(* IEC 61131-3 sources: daoli-st-library/DL_Base (part 4) *)

(* ---- FC_DL_BitCountTransitions.st ---- *)
(*==============================================================================
 * 名称 : FC_DL_BitCountTransitions —— WORD 相邻位跳变统计（总跳变 / 上升 / 下降）
 * 分类 / 前缀 / 版本 : DL_Base / FC_DL_ / 1.0.0
 * 溯源 : 开源语义参考（OSCAT/AixOCAT 族，MIT）或 clean-room IEC 实现，未复制源码
 * 平台 : 纯 IEC 61131-3
 * 功能说明 : 单趟扫描 WORD 的 15 对相邻位（bit i-1 → bit i，i=1..15），统计
 *            跳变总次数并分解为上升（0→1）与下降（1→0）计数；恒有
 *            nRise + nFall = 返回值（调用方可据此自证）。
 *            边界处理：全 0 / 全 1 输入无跳变，三项全 0，属合法结果。
 * 错误码 : 无故障路径（全值域合法的纯统计），eErr 恒 0，bValid 恒 TRUE；
 *          16#0001_1A07 为本件预留码位，当前实现不发出
 * 状态机 : R6 标注 N/A（纯函数无顺序状态，以本节替代 ELSE 兜底）
 * 红线 : R1/R2/R3 ✓ 零全局/零IO/纯IEC ｜ R4 ✓ 移位量≤15 ｜ R10 ✓ 标准转换 ｜ R11 ✓ 分号收尾 ｜ R15 ✓ 无保留字撞名
 * 修订记录 : 2026-11-23 v1.0.0 首次入库（R76）
 *============================================================================*)
FUNCTION FC_DL_BitCountTransitions : INT
VAR_INPUT
    wWord : WORD;      // 待统计的输入字 [位域] / input word to be analyzed
END_VAR
VAR_OUTPUT
    nRise : INT;       // 0→1 上升跳变次数 [次] / number of rising transitions
    nFall : INT;       // 1→0 下降跳变次数 [次] / number of falling transitions
    eErr  : UDINT;     // 故障码，0=正常（本件无故障路径）/ error code, 0=ok (no fault path)
    bError: BOOL;      // 故障标志，恒 FALSE / error flag, always FALSE
    bValid: BOOL;      // TRUE=三项计数可用，恒 TRUE / TRUE when counts are usable
END_VAR
VAR
    _i     : INT;      // 位对扫描游标（取 bit i 与 bit i-1）[位] / pair scan cursor
    _wBit  : WORD;     // 当前位单比特掩码 [位域] / single-bit mask of current bit
    _wPrev : WORD;     // 前一位单比特掩码 [位域] / single-bit mask of previous bit
    _xCur  : BOOL;     // 当前位电平 / level of current bit
    _xPrev : BOOL;     // 前一位电平 / level of previous bit
END_VAR

FC_DL_BitCountTransitions := 0;              // 返回值（总跳变）预设 0 / preset total to zero
nRise := 0;                                  // 上升计数清零 / clear rise count
nFall := 0;                                  // 下降计数清零 / clear fall count
eErr  := 16#0000_0000;                       // 故障码清零 / clear error code
bError:= FALSE;                              // 故障标志清零 / clear error flag
bValid:= TRUE;                               // 本件全值域合法，恒可用 / always valid

FOR _i := 1 TO 15 DO                         // 扫描 15 对相邻位 / scan the 15 adjacent pairs
    _wBit  := SHL(WORD#16#0001, _i);         // 当前位掩码（_i≤15 安全）/ mask of current bit
    _wPrev := SHL(WORD#16#0001, _i - 1);     // 前一位掩码（i-1≥0 安全）/ mask of previous bit
    _xCur  := (wWord AND _wBit)  <> WORD#16#0000;    // 取当前位电平 / sample current bit
    _xPrev := (wWord AND _wPrev) <> WORD#16#0000;    // 取前一位电平 / sample previous bit
    IF _xCur AND (NOT _xPrev) THEN           // 0→1 上升沿 / rising transition
        nRise := nRise + 1;                  // 上升计数加一 / bump rise count
    END_IF
    IF (NOT _xCur) AND _xPrev THEN           // 1→0 下降沿 / falling transition
        nFall := nFall + 1;                  // 下降计数加一 / bump fall count
    END_IF
END_FOR

FC_DL_BitCountTransitions := nRise + nFall;  // 恒等式：总跳变 = 上升 + 下降 / invariant: total = rise + fall

END_FUNCTION

(* ---- FC_DL_BitFieldExtractLword.st ---- *)
(*
  ==================================================================
  组件名 Component  : FC_DL_BitFieldExtractLword
  分类   Category   : DL_Base
  复杂度 Complexity  : 中
  版本   Version    : 1.0.0
  功能   Purpose    : LWORD 单字段提取（起始位 + 宽度 → 右对齐字段值）。全程零
                      64 位移位：先拆高低两个 DWORD 半区，再在半区内做 <=31 位的
                      移位与常量掩码，跨半区时用 DWORD_TO_LWORD 升位拼接。
  来源   Source     : t2-1-lgf-bitlogic（LGF BitLogic 位域提取族 64 位变体）
  溯源   Origin     : 位域提取属公开位运算语义，clean-room 自研实现，未复制 LGF
                      或任何厂商私有库源码。
  平台   Platform   : 纯 IEC 61131-3（AND / OR / SHR / SHL 只作用在 DWORD 域，
                      移位量恒 <32；LWORD 域只出现 AND 与整除），三平台通用
  分工声明 Split     : 与 FC_DL_BitFieldExtract（32 位属主）互引——后者管 DWORD
                      域单字提取；本件为 LWORD 域半区拆分版，不重声明既有位域类型。
  作者   Author     : 道莅代码库 · PLC 编程专家（R60）
  ------------------------------------------------------------------
  边界 Boundary     :
                      一 全程零 64 位移位：高 32 位以「整除 2^32 再 LWORD_TO_DWORD」
                         取得（LWORD 域只做 AND 与整除，不做移位），半区内移位量
                         经 MOD 32 归一后恒在 0..31（R48）；
                      二 宽度 32 的掩码走常量 16#FFFF_FFFF，禁写 SHL(x, 32)；
                      三 非 32 对齐下「宽 64 跨两字」在本实现物理不可达（宽 64 只
                         能起始于位 0），此偏离显式声明：start + width > 64 时主动
                         收窄宽度并置截断信息级码，不静默出半个字段；
                      四 非法域：宽度为 0 或起始位 > 63 判故障级码，输出 0 且 bErr；
                      五 无状态纯函数：局部量一律段 1 显式预置（R254）。
  错误码   Codes    :
    16#0001_0616【故障级】字段域非法（宽度 0 或起始位 >63），输出 0
    16#0001_0617【信息级】字段越出 64 位容器，宽度已收窄（bTrunc 同步置位）
  验收   Acceptance :
    算法已证（脚本）：未跑 ｜ 编译器已证（三平台）：未跑
    V1 src=16#FFFF_FFFF_FFFF_FFFF、start=60、width=4 → 字段 16#F，bTrunc=FALSE
    V2 src=16#1234_5678_9ABC_DEF0、start=28、width=8 → 字段 16#BC（跨半区）
    V3 src 任意、start=62、width=8 → 宽度收窄为 2、bTrunc=TRUE、码 0617
    V4 width=0 → bErr=TRUE、码 0616、字段 0
  修订记录 Revision  :
    2026-11-21  v1.0.0  R60 首版（批 2 · 序号 5）
  ==================================================================
*)
FUNCTION FC_DL_BitFieldExtractLword : LWORD
VAR_INPUT
    uSrc   : LWORD; // 源字 [位串] / the source word
    uStart : UINT;  // 字段起始位号 [位]，合法域 0..63 / the field start bit, legal from zero to sixty three
    uWidth : UINT;  // 字段宽度 [位]，合法域 1..64 / the field width, legal from one to sixty four
END_VAR
VAR_OUTPUT
    bTrunc : BOOL;  // 宽度被收窄（越出容器）[-] / the width was narrowed at the container edge
    bErr   : BOOL;  // 域非法标志 [-] / the illegal domain flag
    eErr   : UDINT; // 错误码，0 = 正常 / the error code, zero is ok
    bError : BOOL;  // 错误标志，eErr 非 0 时为真 / the error flag, true when eErr is nonzero
END_VAR
VAR
    dwLow    : DWORD; // 源字低半区 [位串] / the low half of the source
    dwHigh   : DWORD; // 源字高半区 [位串] / the high half of the source
    dwMask   : DWORD; // 半区内字段掩码 [位串] / the field mask inside a half
    dwMaskHi : DWORD; // 跨半区时高半区剩余宽度掩码 [位串] / the remaining width mask on the high half
    dwPart1  : DWORD; // 跨半区低位片段 [位串] / the low fragment of a cross half field
    dwPart2  : DWORD; // 跨半区高位片段 [位串] / the high fragment of a cross half field
    nStart   : UINT;  // 归一后的起始位号 [位] / the normalised start bit
    nWidth   : UINT;  // 归一（收窄）后的宽度 [位] / the normalised width
    nLowW    : UINT;  // 跨半区时低半区可容纳宽度 [位] / the width the low half can hold
    nShift   : UINT;  // 半区内移位量 [位]，恒 0..31 / the shift amount inside a half, always zero through thirty one
END_VAR
VAR CONSTANT
    DL_BFE_32    : UINT := 32;                      // 半区位宽 [位] / the half width
    DL_BFE_ALL   : DWORD := 16#FFFF_FFFF;           // 32 位全一掩码（禁用 SHL(x, 32)）/ the full thirty two bit mask
    DL_BFE_2P32  : LWORD := 16#0000_0001_0000_0000; // 2 的 32 次幂，用于取高半区（LWORD 域整除，不做移位）/ two to the thirty second, used to take the high half by division
END_VAR

// 段 1｜返回值与错误状态预置安全值（四段式第一段，R45）+ 局部量显式预置（R254）/ segment 1, the preset of the return, the codes and the local guards
FC_DL_BitFieldExtractLword := 16#0000_0000_0000_0000; // 返回值预置零 / preset the return to zero
bTrunc := FALSE; // 截断标志预置假 / preset the truncation flag false
bErr := FALSE; // 域非法标志预置假 / preset the domain fault flag false
eErr := 16#0000_0000; // 错误码预置正常 / preset the code to ok
bError := FALSE; // 错误标志预置假 / preset the error flag false
nStart := 0; // 起始位预置零 / preset the start bit zero
nWidth := 0; // 宽度预置零 / preset the width zero
nLowW := 0; // 低半区宽度预置零 / preset the low half width zero
nShift := 0; // 移位量预置零 / preset the shift amount zero
dwMask := 16#0000_0000; // 掩码预置零 / preset the mask zero
dwMaskHi := 16#0000_0000; // 高位掩码预置零 / preset the high mask zero
dwPart1 := 16#0000_0000; // 低位片段预置零 / preset the low fragment zero
dwPart2 := 16#0000_0000; // 高位片段预置零 / preset the high fragment zero

// 段 2｜域闸（下界早退 + 上界钳位，边界三）/ segment 2, the domain gate with the early return and the narrowing
IF (uWidth < 1) OR (uStart > 63) THEN // 宽度为零或起始位越域 / a zero width or a start beyond the container
    bErr := TRUE; // 置域非法标志 / raise the domain fault flag
    eErr := 16#0001_0616; // 故障级：字段域非法 / fault grade, the field domain is illegal
    bError := TRUE; // 置错误标志（R45 配对）/ raise the error flag, paired with the fault code
    RETURN; // 早退：返回值保持零 / early return with the field zero
END_IF
nStart := uStart; // 域内接管起始位 / take the start bit inside the domain
nWidth := uWidth; // 域内接管宽度 / take the width inside the domain
IF (UINT_TO_UDINT(nStart) + UINT_TO_UDINT(nWidth)) > 64 THEN // 越出 64 位容器 / beyond the sixty four bit container
    nWidth := 64 - nStart; // 主动收窄到容器边界（边界三偏离声明）/ narrow to the container edge with the declared deviation
    bTrunc := TRUE; // 置截断标志 / raise the truncation flag
    eErr := 16#0001_0617; // 信息级：宽度已收窄 / informational, the width narrowed
    bError := TRUE; // 置错误标志 / raise the error flag
END_IF

// 段 3｜半区拆分（零 64 位移位，边界一）：低半区截断取，高半区整除取 / segment 3, the half split with no sixty four bit shift
dwLow := LWORD_TO_DWORD(uSrc); // 低半区：截断取低 32 位 / the low half by truncation
dwHigh := LWORD_TO_DWORD(uSrc / DL_BFE_2P32); // 高半区：整除 2^32 后取低 32 位 / the high half by the division

// 段 4｜字段提取与跨半区拼接（掩码先于移位构造，移位量恒 <32）/ segment 4, the extraction and the cross half splice
IF (nWidth = 32) THEN // 宽 32：常量全一掩码（禁 SHL(x, 32)）/ a full half width uses the constant mask
    dwMask := DL_BFE_ALL; // 常量掩码 / the constant mask
ELSE // 宽 1..31：SHL(1, nWidth) - 1，移位量最大 31 结构性安全 / widths one through thirty one
    dwMask := SHL(DWORD#1, nWidth) - DWORD#1; // 低位起的 nWidth 个一并 / the nWidth low bits set
END_IF
IF nStart >= DL_BFE_32 THEN // 字段整段落在高半区 / the field lies entirely in the high half
    nShift := nStart - DL_BFE_32; // 半区内移位量 0..31 / the shift inside the half, zero through thirty one
    FC_DL_BitFieldExtractLword := DWORD_TO_LWORD(SHR(dwHigh AND dwMask, nShift)); // 高半区提取后升位 / extract from the high half then widen
ELSIF (UINT_TO_UDINT(nStart) + UINT_TO_UDINT(nWidth)) <= 32 THEN // 字段整段落在低半区 / the field lies entirely in the low half
    nShift := nStart; // 半区内移位量 0..31 / the shift inside the half, zero through thirty one
    FC_DL_BitFieldExtractLword := DWORD_TO_LWORD(SHR(dwLow AND dwMask, nShift)); // 低半区提取后升位 / extract from the low half then widen
ELSE // 跨半区：低片段 + 高片段移位拼接（nStart 必在 1..31）/ a cross half field, both fragments spliced
    nLowW := 32 - nStart; // 低半区可容纳宽度 1..31 / the width the low half holds, one through thirty one
    IF nLowW >= 32 THEN // 结构性不可达（nStart ≥ 1 恒真），显式兜底防掩码移位越界 / structurally unreachable, kept as an explicit guard
        nLowW := 31; // 兜底收窄到 31 位 / narrow to thirty one bits
    END_IF
    dwPart1 := SHR(dwLow AND (SHL(DWORD#1, nLowW) - DWORD#1), nStart); // 低片段右移到最低位 / shift the low fragment down to bit zero
    dwMaskHi := SHL(DWORD#1, nWidth - nLowW) - DWORD#1; // 高半区剩余宽度掩码 / the remaining width mask on the high half
    dwPart2 := SHL(dwHigh AND dwMaskHi, nLowW); // 高片段左移到低片段之上（移位量 1..31）/ shift the high fragment above the low one
    FC_DL_BitFieldExtractLword := DWORD_TO_LWORD(dwPart1 OR dwPart2); // 两片段拼合后升位 / splice then widen
END_IF

// 段 5｜结果复检：字段宽度上界自证（nWidth ≤ 64，拼接已按半区完成，无溢出路径）/ segment 5, the result recheck
IF bTrunc AND (nWidth >= 1) THEN // 收窄后仍为合法宽度 / the narrowed width is still legal
    eErr := 16#0001_0617; // 信息级：宽度已收窄（回放，防段 4 覆盖）/ informational, the width narrowed, replayed against the overwrite
END_IF
END_FUNCTION

(* ---- FC_DL_BitFillLowestZero.st ---- *)
(*==============================================================================
 * 名称 : FC_DL_BitFillLowestZero —— 最低 0 位置 1（DWORD），输出该位位号
 * 分类 / 前缀 / 版本 : DL_Base / FC_DL_ / 1.0.0
 * 溯源 : 开源语义参考（OSCAT/AixOCAT 族，MIT）或 clean-room IEC 实现，未复制源码
 * 平台 : 纯 IEC 61131-3
 * 功能说明 : 把输入 DWORD 中最低的 0 位置 1 后返回（即 dwIn OR 单比特隔离值），
 *            并给出该位位号 nPos。常用于资源位图分配（找空位并占用）。
 *            边界处理：输入全 1 时无 0 位可填，原值返回、nPos=-1、bValid=FALSE
 *            并置 eErr（返回值虽为原值，但语义上未发生分配）。
 * 错误码 : 16#0001_1A08 = 输入全 1，无 0 位可填
 *          eErr=0 且 bValid=TRUE 表示已完成填位且 nPos 有效
 * 状态机 : R6 标注 N/A（纯函数无顺序状态，以本节替代 ELSE 兜底）
 * 红线 : R1/R2/R3 ✓ 零全局/零IO/纯IEC ｜ R4 ✓ 移位量≤31 ｜ R10 ✓ 标准转换 ｜ R11 ✓ 分号收尾 ｜ R15 ✓ 无保留字撞名
 * 修订记录 : 2026-11-23 v1.0.0 首次入库（R76）
 *============================================================================*)
FUNCTION FC_DL_BitFillLowestZero : DWORD
VAR_INPUT
    dwIn : DWORD;      // 输入位图 [位域] / input bitmap dword
END_VAR
VAR_OUTPUT
    nPos   : INT;      // 被填 1 的最低 0 位位号，全 1 时为 -1 [位] / bit index filled, -1 if none
    eErr   : UDINT;    // 故障码，0=正常，1A08=全 1 无空位 / error code, 0=ok, 1A08=all-ones input
    bError : BOOL;     // TRUE=本件发生故障 / TRUE when fault occurred
    bValid : BOOL;     // TRUE=填位成功且 nPos 有效 / TRUE when fill succeeded and nPos valid
END_VAR
VAR
    _dwNot  : DWORD;   // 输入按位取反（0 位变 1 位）/ inverted input (zeros become ones)
    _dwIso  : DWORD;   // 最低 0 位的单比特隔离值 [位域] / isolated lowest zero bit
    _i      : INT;     // 位扫描游标 [位] / bit scan cursor
    _dwW    : DWORD;   // 单比特游走值 [位域] / single-bit walker
    _xHit   : BOOL;    // 命中标志 / found flag
END_VAR

nPos := -1;                                  // 位号预设 -1（未命中语义）/ preset position to -1
eErr   := 16#0000_0000;                      // 故障码清零 / clear error code
bError := FALSE;                             // 故障标志清零 / clear error flag
bValid := TRUE;                              // 预设输出可用 / preset valid flag

_dwNot := NOT dwIn;                          // 取反后 0 位变 1 位 / invert so zeros become ones
IF _dwNot = DWORD#16#0000_0000 THEN          // 全 1：无 0 位可填 / all ones: nothing to fill
    eErr   := 16#0001_1A08;                  // 置全 1 故障码 / set all-ones code
    bError := TRUE;                          // 置故障标志 / set error flag
    bValid := FALSE;                         // nPos 不可用 / position not usable
    FC_DL_BitFillLowestZero := dwIn;         // 原值返回 / return input unchanged
    RETURN;                                  // 提前收口 / early exit
END_IF

_dwIso := _dwNot AND (NOT (_dwNot - DWORD#16#0000_0001));    // 隔离最低 0 位（同最低 1 位法）/ isolate lowest zero bit
_xHit  := FALSE;                             // 命中标志清零 / clear found flag
FOR _i := 0 TO 31 DO                         // 从低位找第一个命中 / scan low to high for first hit
    _dwW := SHL(DWORD#16#0000_0001, _i);     // 当前位单比特掩码（_i≤31 安全）/ single-bit mask
    IF (NOT _xHit) AND ((_dwIso AND _dwW) <> DWORD#16#0000_0000) THEN    // 首个命中即停扫 / stop at first hit
        nPos  := _i;                         // 回写位号 / write back bit index
        _xHit := TRUE;                       // 置命中标志 / set found flag
    END_IF
END_FOR

FC_DL_BitFillLowestZero := dwIn OR _dwIso;   // 填 1 后返回 / return with the bit filled

END_FUNCTION

(* ---- FC_DL_BitGet.st ---- *)
(*==============================================================================
 * 组件名称 (Component)  : FC_DL_BitGet
 * 所属子库 (Sublibrary) : DL_Base
 * 当前版本 (Version)    : 1.0.0
 * 兼容性   (Platform)   : CODESYS 3.5 / TwinCAT 3 / 汇川 InoProShop / Machine Expert
 *                         仅用标准 SHR / AND 运算，无任何厂商位访问语法
 * 功能描述 (Function)   : 从 32 位状态字中安全提取指定位（Hamming 单位提取）。
 *                         位索引合法域 0..31（0 = LSB）。越界时"先判后算"，
 *                         立即返回 FALSE 并输出 16#0001_0001，绝不把越界移位量
 *                         交给 SHL/SHR 去执行（越界移位在各平台行为不一致，是
 *                         跨平台移植的经典暗坑）。
 * 开源溯源 (Origin)     : 原创实现。位序约定遵循 IEC 61131-3 对位串类型
 *                         "第 0 位为最低有效位"的规定。
 * 依赖     (Depends)    : 无 DL_ 内部依赖；无标准库功能块依赖
 * 红线自检 (Redline)    : R1 ✓ 零全局变量表与外部变量引用 ｜ R2 ✓ 零物理 IO 地址直写
 *                         R3 ✓ 纯 IEC 61131-3（无厂商位访问方言）｜ R4 ✓ 越界先判后算 + 返回值兜底
 *                         R5 ✓ 全变量中英双语同行注释 ｜ R6 N/A（无状态机）｜ R7 N/A（无实例调用）
 * 修订历史 (Revision)   :
 *   2026-11-14  v1.0.0  首版入库（Phase 1 冷启动 · Level 0 批次）
 *============================================================================*)
FUNCTION FC_DL_BitGet : BOOL
VAR_INPUT
    uValue    : DWORD;    // 待检测的 32 位状态字 / Source 32-bit status word
    uBitIndex : USINT;    // 位序号，0 = LSB，合法域 0..31 / Bit index, 0 = LSB, valid range 0..31
END_VAR
VAR_OUTPUT
    bValid    : BOOL;     // 索引合法标志，FALSE 时返回值为保底 FALSE / Index valid flag, FALSE means result is a safe FALSE
    uErrorId  : UDINT;    // 故障码，0 = 无故障 / Error code, 0 = no error
END_VAR
VAR
    uWork     : UDINT;    // 提升到 UDINT 的工作副本，规避混合类型移位 / UDINT working copy to avoid mixed-type shifts
    uShift    : UDINT;    // 提升到 UDINT 的移位量 / Shift amount promoted to UDINT
END_VAR
VAR CONSTANT
    DL_BIT_INDEX_MAX : USINT := 31;  // 32 位字的最大合法位索引 / Max legal bit index of a 32-bit word
END_VAR

(*------------------------------------------------------------------------------
 * 段 1｜返回值与标志预置：任何异常路径下返回值必须确定
 *      Pre-set return value and flags: the result must be deterministic on every path
 *      部分平台函数返回值未赋值时残留上次调用值，故先给 FALSE（边界 B4）
 *-----------------------------------------------------------------------------*)
FC_DL_BitGet := FALSE;
bValid       := FALSE;
uErrorId     := 16#0000_0000;
uWork        := 16#0000_0000;

(*------------------------------------------------------------------------------
 * 段 2｜越界先判后算（边界 B1）：禁止先移位再校验
 *      Bounds check before any shift (boundary B1): never shift first and check later
 *      USINT 全域 0..255，凡 > 31 者均属非法移位量，统一按参数越界处理
 *-----------------------------------------------------------------------------*)
IF uBitIndex > DL_BIT_INDEX_MAX THEN
    uErrorId := 16#0001_0001;
    RETURN;
END_IF

(*------------------------------------------------------------------------------
 * 段 3｜位提取（边界 B2/B3）：统一提升到 UDINT 后移位，再显式掩码取最低位
 *      Bit extraction: promote to UDINT, shift, then mask the LSB explicitly
 *      禁止使用以点号直取单一位的厂商方言；禁止依赖"非零即真"的隐式布尔转换
 *-----------------------------------------------------------------------------*)
uWork  := DWORD_TO_UDINT(uValue);
uShift := USINT_TO_UDINT(uBitIndex);
uWork  := SHR(uWork, uShift);
uWork  := uWork AND 16#0000_0001;

IF uWork <> 16#0000_0000 THEN
    FC_DL_BitGet := TRUE;
END_IF

(* 校验通过：索引合法，结果可信 *)
(* Check passed: index is legal and the result is trustworthy *)
bValid := TRUE;
END_FUNCTION

(* ---- FC_DL_BitLowestSet.st ---- *)
(*==============================================================================
 * 名称 : FC_DL_BitLowestSet —— 最低置位位号与单比特隔离值（DWORD）
 * 分类 / 前缀 / 版本 : DL_Base / FC_DL_ / 1.0.0
 * 溯源 : 开源语义参考（OSCAT/AixOCAT 族，MIT）或 clean-room IEC 实现，未复制源码
 * 平台 : 纯 IEC 61131-3
 * 功能说明 : 返回输入 DWORD 中最低置位位的位号（0..31），并输出单比特隔离值
 *            dwIsolate = dwIn AND (NOT (dwIn - 1))（无符号回绕语义，等价于
 *            二进制补码的 x AND (-x)，仅保留最低的 1 位）。
 *            边界处理：dwIn 全 0 时无置位位，返回 -1、dwIsolate=0、bValid=FALSE
 *            并置 eErr（隔离值无效，调用方不得使用）。
 * 错误码 : 16#0001_1A05 = 输入全 0，无置位位可隔离
 *          eErr=0 且 bValid=TRUE 表示返回位号与隔离值均有效
 * 状态机 : R6 标注 N/A（纯函数无顺序状态，以本节替代 ELSE 兜底）
 * 红线 : R1/R2/R3 ✓ 零全局/零IO/纯IEC ｜ R4 ✓ 移位量≤31 ｜ R10 ✓ 标准转换 ｜ R11 ✓ 分号收尾 ｜ R15 ✓ 无保留字撞名
 * 修订记录 : 2026-11-23 v1.0.0 首次入库（R76）
 *============================================================================*)
FUNCTION FC_DL_BitLowestSet : INT
VAR_INPUT
    dwIn : DWORD;      // 待扫描的输入双字 [位域] / input dword to be scanned
END_VAR
VAR_OUTPUT
    dwIsolate : DWORD;    // 最低置位位的单比特隔离值 [位域] / isolated lowest set bit
    eErr      : UDINT;    // 故障码，0=正常，1A05=输入全 0 / error code, 0=ok, 1A05=all-zero input
    bError    : BOOL;     // TRUE=本件发生故障 / TRUE when fault occurred
    bValid    : BOOL;     // TRUE=返回位号与隔离值可用 / TRUE when outputs are usable
END_VAR
VAR
    _i    : INT;       // 位扫描游标 [位] / bit scan cursor
    _dwW  : DWORD;     // 单比特游走值 [位域] / single-bit walker
    _xHit : BOOL;      // 是否已找到最低置位位 / found flag for lowest set bit
END_VAR

FC_DL_BitLowestSet := -1;                    // 返回值预设 -1（未命中语义）/ preset return to -1
dwIsolate := DWORD#16#0000_0000;             // 隔离值预设全 0 / preset isolate to zero
eErr      := 16#0000_0000;                   // 故障码清零 / clear error code
bError    := FALSE;                          // 故障标志清零 / clear error flag
bValid    := TRUE;                           // 预设输出可用 / preset valid flag

IF dwIn = DWORD#16#0000_0000 THEN            // 输入全 0：无置位位 / all-zero input: no set bit
    eErr   := 16#0001_1A05;                  // 置全 0 故障码 / set all-zero code
    bError := TRUE;                          // 置故障标志 / set error flag
    bValid := FALSE;                         // 位号与隔离值均不可用 / outputs not usable
    RETURN;                                  // 返回 -1、隔离值 0 / return -1 with zero isolate
END_IF

dwIsolate := dwIn AND (NOT (dwIn - DWORD#16#0000_0001));    // 经典隔离式，仅留最低 1 位 / classic isolate of lowest set bit
_xHit := FALSE;                              // 命中标志清零 / clear found flag
FOR _i := 0 TO 31 DO                         // 从低位向高位找第一个 1 / scan low to high for first one
    _dwW := SHL(DWORD#16#0000_0001, _i);     // 当前位单比特掩码（_i≤31 安全）/ single-bit mask
    IF (NOT _xHit) AND ((dwIsolate AND _dwW) <> DWORD#16#0000_0000) THEN    // 首个命中即停扫 / stop at first hit
        FC_DL_BitLowestSet := _i;            // 回写最低置位位号 / write back lowest bit index
        _xHit := TRUE;                       // 置命中标志 / set found flag
    END_IF
END_FOR

END_FUNCTION

(* ---- FC_DL_BitMaskRange.st ---- *)
(*==============================================================================
 * 名称 : FC_DL_BitMaskRange —— 连续位区间掩码构造（bitLo..bitHi 置 1 的 DWORD 掩码）
 * 分类 / 前缀 / 版本 : DL_Base / FC_DL_ / 1.0.0
 * 溯源 : 开源语义参考（OSCAT/AixOCAT 族，MIT）或 clean-room IEC 实现，未复制源码
 * 平台 : 纯 IEC 61131-3
 * 功能说明 : 依入参位号 uLo..uHi 构造 DWORD 掩码，区间内各位置 1、其余为 0。
 *            边界处理：uLo/uHi 越界（<0 或 >31）先钳位到 [0,31] 再构造；
 *            钳位后 uLo>uHi（区间为空）返回 DWORD#0 并置 eErr 故障码。
 *            移位量恒 ≤31（<DWORD 位宽 32），结构性无越界移位。
 * 错误码 : 16#0001_1A01 = 钳位后位区间为空（uLo>uHi），掩码无意义
 *          eErr=0 且 bValid=TRUE 表示掩码有效；bValid=FALSE 时返回值勿用
 * 状态机 : R6 标注 N/A（纯函数无顺序状态，以本节替代 ELSE 兜底）
 * 红线 : R1/R2/R3 ✓ 零全局/零IO/纯IEC ｜ R4 ✓ 移位量≤31 ｜ R10 ✓ 标准转换 ｜ R11 ✓ 分号收尾 ｜ R15 ✓ 无保留字撞名
 * 修订记录 : 2026-11-23 v1.0.0 首次入库（R76）
 *============================================================================*)
FUNCTION FC_DL_BitMaskRange : DWORD
VAR_INPUT
    uLo : INT;     // 起始位号 0..31，越界自动钳位 [位] / low bit index, clamped into [0,31]
    uHi : INT;     // 结束位号 0..31，越界自动钳位 [位] / high bit index, clamped into [0,31]
END_VAR
VAR_OUTPUT
    eErr   : UDINT;    // 故障码，0=正常，1A01=区间为空 / error code, 0=ok, 1A01=empty range
    bError : BOOL;     // TRUE=本件发生参数级故障 / TRUE when parameter-level fault occurred
    bValid : BOOL;     // TRUE=返回值可用 / TRUE when return value is usable
END_VAR
VAR
    _nLo   : INT;      // 钳位后的起始位号 [位] / clamped low bit index
    _nHi   : INT;      // 钳位后的结束位号 [位] / clamped high bit index
    _i     : INT;      // 位扫描游标 [位] / bit scan cursor
    _dwBit : DWORD;    // 当前游标对应的单比特值 [位域] / single-bit walker value
END_VAR

FC_DL_BitMaskRange := DWORD#16#0000_0000;    // 返回值预设全 0 掩码 / preset return to zero mask
eErr   := 16#0000_0000;                      // 故障码清零 / clear error code
bError := FALSE;                             // 故障标志清零 / clear error flag
bValid := TRUE;                              // 预设输出可用 / preset valid flag

_nLo := uLo;                                 // 取入参起始位号 / take input low index
_nHi := uHi;                                 // 取入参结束位号 / take input high index
IF _nLo < 0 THEN _nLo := 0; END_IF           // 下界钳位 / clamp lower bound
IF _nLo > 31 THEN _nLo := 31; END_IF         // 上界钳位 / clamp upper bound
IF _nHi < 0 THEN _nHi := 0; END_IF           // 下界钳位 / clamp lower bound
IF _nHi > 31 THEN _nHi := 31; END_IF         // 上界钳位 / clamp upper bound

IF _nLo > _nHi THEN                          // 钳位后区间为空 / empty range after clamping
    eErr   := 16#0001_1A01;                  // 置区间为空故障码 / set empty-range code
    bError := TRUE;                          // 置故障标志 / set error flag
    bValid := FALSE;                         // 返回值不可用 / return value not usable
    RETURN;                                  // 返回值保持全 0 掩码 / return stays zero mask
END_IF

_dwBit := SHL(DWORD#16#0000_0001, _nLo);     // 单比特走到起始位（_nLo≤31 安全）/ walk bit to start
FOR _i := _nLo TO _nHi DO                    // 逐位置 1 / set bits one by one
    FC_DL_BitMaskRange := FC_DL_BitMaskRange OR _dwBit;    // 并入当前位 / merge current bit
    _dwBit := SHL(_dwBit, 1);                // 单比特左移一位，循环内 _i<_nHi≤31 安全 / shift walker left
END_FOR

END_FUNCTION

(* ---- FC_DL_BitReverse16.st ---- *)
(*==============================================================================
 * 名称 : FC_DL_BitReverse16 —— WORD 位序完全反转（bit0↔bit15 镜像）
 * 分类 / 前缀 / 版本 : DL_Base / FC_DL_ / 1.0.0
 * 溯源 : 开源语义参考（OSCAT/AixOCAT 族，MIT）或 clean-room IEC 实现，未复制源码
 * 平台 : 纯 IEC 61131-3
 * 功能说明 : 将 WORD 的 16 个位按镜像序重排后返回（第 i 位映射到第 15-i 位）。
 *            边界处理：全 0 / 全 1 / 回文位型（如 16#8081）均原值返回，属合法结果；
 *            循环固定 16 次，无越界移位（i 与 15-i 均 ≤15 < 16 位宽）。
 * 错误码 : 无故障路径（全值域合法的纯变换），eErr 恒 0，bValid 恒 TRUE；
 *          16#0001_1A03 为本件预留码位，当前实现不发出
 * 状态机 : R6 标注 N/A（纯函数无顺序状态，以本节替代 ELSE 兜底）
 * 红线 : R1/R2/R3 ✓ 零全局/零IO/纯IEC ｜ R4 ✓ 移位量≤15 ｜ R10 ✓ 标准转换 ｜ R11 ✓ 分号收尾 ｜ R15 ✓ 无保留字撞名
 * 修订记录 : 2026-11-23 v1.0.0 首次入库（R76）
 *============================================================================*)
FUNCTION FC_DL_BitReverse16 : WORD
VAR_INPUT
    wIn : WORD;        // 待反转的输入字 [位域] / input word to be bit-reversed
END_VAR
VAR_OUTPUT
    eErr   : UDINT;    // 故障码，0=正常（本件无故障路径）/ error code, 0=ok (no fault path)
    bError : BOOL;     // 故障标志，恒 FALSE / error flag, always FALSE
    bValid : BOOL;     // TRUE=返回值可用，恒 TRUE / TRUE when return value is usable
END_VAR
VAR
    _i     : INT;      // 位扫描游标 [位] / bit scan cursor
    _wBit  : WORD;     // 当前读出位对应的单比特值 [位域] / single-bit walker for read side
END_VAR

FC_DL_BitReverse16 := WORD#16#0000;          // 返回值预设全 0 / preset return to zero
eErr   := 16#0000_0000;                      // 故障码清零 / clear error code
bError := FALSE;                             // 故障标志清零 / clear error flag
bValid := TRUE;                              // 本件全值域合法，恒可用 / always valid

FOR _i := 0 TO 15 DO                         // 逐位镜像搬运 / mirror bits one by one
    _wBit := SHL(WORD#16#0001, _i);          // 读侧单比特（_i≤15 安全）/ single bit on read side
    IF (wIn AND _wBit) <> WORD#16#0000 THEN  // 源位为 1 才搬运 / copy only when source bit set
        FC_DL_BitReverse16 := FC_DL_BitReverse16 OR SHL(WORD#16#0001, 15 - _i);    // 写入镜像位（15-_i≤15 安全）/ set mirrored bit
    END_IF
END_FOR

END_FUNCTION

(* ---- FC_DL_BitReverse8.st ---- *)
(*==============================================================================
 * 名称 : FC_DL_BitReverse8 —— BYTE 位序完全反转（bit0↔bit7 镜像）
 * 分类 / 前缀 / 版本 : DL_Base / FC_DL_ / 1.0.0
 * 溯源 : 开源语义参考（OSCAT/AixOCAT 族，MIT）或 clean-room IEC 实现，未复制源码
 * 平台 : 纯 IEC 61131-3
 * 功能说明 : 将 BYTE 的 8 个位按镜像序重排后返回（第 i 位映射到第 7-i 位）。
 *            边界处理：全 0 / 全 1 / 回文位型（如 16#18）均原值返回，属合法结果；
 *            循环固定 8 次，无越界移位（i 与 7-i 均 ≤7 < 8 位宽）。
 * 错误码 : 无故障路径（全值域合法的纯变换），eErr 恒 0，bValid 恒 TRUE；
 *          16#0001_1A02 为本件预留码位，当前实现不发出
 * 状态机 : R6 标注 N/A（纯函数无顺序状态，以本节替代 ELSE 兜底）
 * 红线 : R1/R2/R3 ✓ 零全局/零IO/纯IEC ｜ R4 ✓ 移位量≤7 ｜ R10 ✓ 标准转换 ｜ R11 ✓ 分号收尾 ｜ R15 ✓ 无保留字撞名
 * 修订记录 : 2026-11-23 v1.0.0 首次入库（R76）
 *============================================================================*)
FUNCTION FC_DL_BitReverse8 : BYTE
VAR_INPUT
    byIn : BYTE;       // 待反转的输入字节 [位域] / input byte to be bit-reversed
END_VAR
VAR_OUTPUT
    eErr   : UDINT;    // 故障码，0=正常（本件无故障路径）/ error code, 0=ok (no fault path)
    bError : BOOL;     // 故障标志，恒 FALSE / error flag, always FALSE
    bValid : BOOL;     // TRUE=返回值可用，恒 TRUE / TRUE when return value is usable
END_VAR
VAR
    _i     : INT;      // 位扫描游标 [位] / bit scan cursor
    _dwBit : BYTE;     // 当前读出位对应的单比特值 [位域] / single-bit walker for read side
END_VAR

FC_DL_BitReverse8 := BYTE#16#00;             // 返回值预设全 0 / preset return to zero
eErr   := 16#0000_0000;                      // 故障码清零 / clear error code
bError := FALSE;                             // 故障标志清零 / clear error flag
bValid := TRUE;                              // 本件全值域合法，恒可用 / always valid

FOR _i := 0 TO 7 DO                          // 逐位镜像搬运 / mirror bits one by one
    _dwBit := SHL(BYTE#16#01, _i);           // 读侧单比特（_i≤7 安全）/ single bit on read side
    IF (byIn AND _dwBit) <> BYTE#16#00 THEN  // 源位为 1 才搬运 / copy only when source bit set
        FC_DL_BitReverse8 := FC_DL_BitReverse8 OR SHL(BYTE#16#01, 7 - _i);    // 写入镜像位（7-_i≤7 安全）/ set mirrored bit
    END_IF
END_FOR

END_FUNCTION

(* ---- FC_DL_BitRunLength.st ---- *)
(*==============================================================================
 * 名称 : FC_DL_BitRunLength —— WORD 最长连续 1 游程长度与起始位号
 * 分类 / 前缀 / 版本 : DL_Base / FC_DL_ / 1.0.0
 * 溯源 : 开源语义参考（OSCAT/AixOCAT 族，MIT）或 clean-room IEC 实现，未复制源码
 * 平台 : 纯 IEC 61131-3
 * 功能说明 : 单趟扫描 WORD 的 16 个位，返回最长连续 1 的游程长度（0..16），
 *            并给出该游程的起始位号 nStart（0..15）。多条等长游程取最低起始位。
 *            边界处理：无任何 1 位时返回 0 且 nStart=-1（合法结果，非故障，
 *            bValid 保持 TRUE）；游程到字尾截断同样按已计长度参与比较。
 * 错误码 : 无故障路径（全值域合法的纯统计），eErr 恒 0，bValid 恒 TRUE；
 *          16#0001_1A04 为本件预留码位，当前实现不发出
 * 状态机 : R6 标注 N/A（纯函数无顺序状态，以本节替代 ELSE 兜底）
 * 红线 : R1/R2/R3 ✓ 零全局/零IO/纯IEC ｜ R4 ✓ 移位量≤15 ｜ R10 ✓ 标准转换 ｜ R11 ✓ 分号收尾 ｜ R15 ✓ 无保留字撞名
 * 修订记录 : 2026-11-23 v1.0.0 首次入库（R76）
 *============================================================================*)
FUNCTION FC_DL_BitRunLength : INT
VAR_INPUT
    wWord : WORD;      // 待扫描的输入字 [位域] / input word to be scanned
END_VAR
VAR_OUTPUT
    nStart : INT;      // 最长游程起始位号，无 1 时为 -1 [位] / start bit of longest run, -1 if none
    eErr   : UDINT;    // 故障码，0=正常（本件无故障路径）/ error code, 0=ok (no fault path)
    bError : BOOL;     // 故障标志，恒 FALSE / error flag, always FALSE
    bValid : BOOL;     // TRUE=返回值可用，恒 TRUE / TRUE when return value is usable
END_VAR
VAR
    _i        : INT;       // 位扫描游标 [位] / bit scan cursor
    _nCur     : INT;       // 当前游程长度 [位] / current run length
    _nCurSt   : INT;       // 当前游程起始位号 [位] / current run start bit
    _nBest    : INT;       // 已发现的最长游程长度 [位] / best run length so far
    _nBestSt  : INT;       // 已发现的最长游程起始位号 [位] / best run start bit so far
    _wBit     : WORD;      // 当前位单比特掩码 [位域] / single-bit mask of current position
    _xBit     : BOOL;      // 当前位电平 / level of current bit
END_VAR

FC_DL_BitRunLength := 0;                     // 返回值预设 0 / preset return to zero
nStart := -1;                                // 起始位预设 -1（无 1 语义）/ preset start to -1
eErr   := 16#0000_0000;                      // 故障码清零 / clear error code
bError := FALSE;                             // 故障标志清零 / clear error flag
bValid := TRUE;                              // 本件全值域合法，恒可用 / always valid

_nBest  := 0;                                // 最长游程清零 / clear best length
_nBestSt := -1;                              // 最长游程起始清零 / clear best start
_nCur   := 0;                                // 当前游程清零 / clear current length
_nCurSt := 0;                                // 当前游程起始清零 / clear current start

FOR _i := 0 TO 15 DO                         // 单趟从低位到高位扫描 / single low-to-high pass
    _wBit := SHL(WORD#16#0001, _i);          // 当前位单比特掩码（_i≤15 安全）/ single-bit mask
    _xBit := (wWord AND _wBit) <> WORD#16#0000;    // 取当前位电平 / sample current bit
    IF _xBit THEN                            // 位为 1：游程延续或新开 / bit set: extend or open run
        IF _nCur = 0 THEN
            _nCurSt := _i;                   // 新游程序幕，记起始位 / new run starts here
        END_IF
        _nCur := _nCur + 1;                  // 游程长度加一 / extend run length
        IF _nCur > _nBest THEN               // 严格大于保证等长取最低起始位 / strict gt keeps lowest start on ties
            _nBest   := _nCur;               // 刷新最长游程 / refresh best length
            _nBestSt := _nCurSt;             // 刷新最长游程起始位 / refresh best start bit
        END_IF
    ELSE                                     // 位为 0：当前游程终结 / bit clear: current run ends
        _nCur := 0;                          // 游程长度归零 / reset current length
    END_IF
END_FOR

FC_DL_BitRunLength := _nBest;                // 回写最长游程长度 / write back best length
nStart := _nBestSt;                          // 回写起始位号（无 1 时保持 -1）/ write back start bit

END_FUNCTION

(* ---- FC_DL_BitScanLword.st ---- *)
(*
  ==================================================================
  组件名 Component  : FC_DL_BitScanLword
  分类   Category   : DL_Base
  前缀   Naming     : FC_DL_ ｜ b/n/u/f/t/e/st 类型前缀制（R265）
  复杂度 Complexity  : 低
  版本   Version    : 1.0.0
  功能   Purpose    : LWORD 最低/最高置位索引扫描（uIdx + bFound 双出口）。
  来源   Source     : self-std（IEC 标准位操作语义自研包装）
  平台   Platform   : 纯 IEC 61131-3（FOR / AND / SHR / SHL / 比较），三平台通用
  分工声明 Split     : 与 FC_DL_ReverseBitsLword（位序反转属主）分工——本件只做
                      置位索引定位，不改位序；方向由 bHighFirst 选择，不设两个 POU。
  作者   Author     : 道莅代码库 · PLC 编程专家（R61）
  归属 Ownership     : 本件无 TYPE 声明；引用件类型全部 IEC 标准原生。
  ------------------------------------------------------------------
  边界 Boundary     :
                      一 全零输入：bFound = FALSE 且 uIdx = 0（不泄 -1，不泄哨兵），
                         置信息级码（R90 反证：bFound 只表达「有命中」，无法区分
                         「扫描过且全零」与「未扫」，码位补足该可观测性）；
                      二 扫描循环有界恰好 64 次（禁 WHILE 裸循环，防死锁纪律）；
                      三 方向选择：bHighFirst = FALSE 自低位向高位扫（首命中即
                         最低置位），TRUE 自高位向低位扫（首命中即最高置位）；
                      四 无状态纯函数：局部量段 1 显式预置（R254）。
  错误码   Codes    :
    16#0001_0641【信息级】全零输入零命中（bFound = FALSE，uIdx = 0）
  验收   Acceptance :
    算法已证（脚本）：未跑 ｜ 编译器已证（三平台）：未跑
    V1 uSrc=16#0000_0000_0000_0100、bHighFirst=FALSE → uIdx=8、bFound=TRUE
    V2 uSrc=16#0000_0000_0000_0100、bHighFirst=TRUE → uIdx=8（单置位两向同值）
    V3 uSrc=16#0000_0000_0000_0105、bHighFirst=TRUE → uIdx=8
    V4 uSrc=0 → bFound=FALSE、uIdx=0、码 0641
  修订记录 Revision  :
    2026-11-21  v1.0.0  R61 首版（批 1 · 序号 2）
  ==================================================================
*)
FUNCTION FC_DL_BitScanLword : BOOL
VAR_IN_OUT
    uSrc : LWORD; // 待扫描源字 [位图] / the source word to scan
END_VAR
VAR_INPUT
    bHighFirst : BOOL; // 方向开关：TRUE 自高位向低位扫 / the direction switch, true scans from the high end
END_VAR
VAR_OUTPUT
    uIdx   : UDINT; // 首命中置位索引 [位]，零命中时为 0 / the first hit bit index, zero on a miss
    bFound : BOOL;  // 是否存在置位位 [-] / the hit flag
    bValid : BOOL;  // 扫描完成标志（恒真：扫描全域有界）[-] / the scan done flag, always true
    eErr   : UDINT; // 错误码，0 = 正常 / the error code, zero is ok
    bError : BOOL;  // 错误标志（信息级不置位，R285 口径）/ the error flag, never raised by the informational grade
END_VAR
VAR
    k : DINT; // 位循环索引 [位] / the bit loop index
END_VAR

// 段 1｜返回值与输出预置（局部量显式预置，R254）/ segment 1, the preset
FC_DL_BitScanLword := FALSE; // 返回值预置假 / preset the return false
uIdx := 0; // 索引预置零（零命中口径，边界一）/ preset the index zero
bFound := FALSE; // 命中标志预置假 / preset the hit flag false
bValid := FALSE; // 完成标志预置假（出口置真）/ preset the done flag false
eErr := 16#0000_0000; // 错误码预置正常 / preset the code to ok
bError := FALSE; // 错误标志预置假 / preset the error flag false

IF uSrc = 16#0000_0000_0000_0000 THEN // 全零输入：零命中早出（边界一）/ the all zero source, a miss with the declared code
    eErr := 16#0001_0641; // 信息级：零命中（信息级不置 bError）/ informational, the miss without the fault bit
    bValid := TRUE; // 扫描完成 / the scan is done
    FC_DL_BitScanLword := TRUE; // 返回成功 / return success
    RETURN; // 早退 / early return
END_IF

// 段 2｜有界扫描：恰好 64 次，首命中即记（边界二）/ segment 2, the bounded scan of exactly sixty four rounds
IF NOT bHighFirst THEN // 自低位向高位 / from the low end
    FOR k := 0 TO 63 DO // 有界循环 / the bounded loop
        IF NOT bFound THEN // 尚未命中才继续判（首命中口径）/ judge only before the first hit
            IF (uSrc AND SHL(16#0000_0000_0000_0001, k)) <> 16#0000_0000_0000_0000 THEN // 第 k 位为置位 / the bit k is set
                uIdx := DINT_TO_UDINT(k); // 记录命中索引 / register the hit index
                bFound := TRUE; // 置命中标志 / raise the hit flag
            END_IF
        END_IF
    END_FOR
ELSE // 自高位向低位 / from the high end
    FOR k := 63 TO 0 BY -1 DO // 有界反序循环 / the bounded reverse loop
        IF NOT bFound THEN // 尚未命中才继续判 / judge only before the first hit
            IF (uSrc AND SHL(16#0000_0000_0000_0001, k)) <> 16#0000_0000_0000_0000 THEN // 第 k 位为置位 / the bit k is set
                uIdx := DINT_TO_UDINT(k); // 记录命中索引 / register the hit index
                bFound := TRUE; // 置命中标志 / raise the hit flag
            END_IF
        END_IF
    END_FOR
END_IF

// 段 3｜出口（源字非零已证，bFound 必为真）/ segment 3, the outlet, the hit is proven since the source is nonzero
bValid := TRUE; // 扫描完成 / the scan is done
FC_DL_BitScanLword := TRUE; // 返回成功 / return success
END_FUNCTION

(* ---- FC_DL_BitSegmentBlockMove.st ---- *)
(*
    FC_DL_BitSegmentBlockMove —— 跨字多段位段一次搬运
    ------------------------------------------------------------------
    分类      : DL_Base / BitString
    前缀      : FC_DL_
    版本      : 1.0.0
    溯源      : T2-1 LGF · Bit Logic（只借「读 / 写 / 监视 三层粒度 + 批量段」的组内
                分类事实；库内已收口 Extract / Insert / ChangeWatch 三件，本件补
                「多段一次搬」缺口）；掩码、段表结构、判界顺序、码位 100% 自有；
                clean-room 重写，未复制任何闭源厂商源码，参考实现仅限 MIT/Apache 许可
    平台      : 纯 IEC 61131-3，CODESYS V3.5+ / TwinCAT 3 / InoProShop 通用
    作者      : 道莅代码库 · PLC编程专家（R18）
    ------------------------------------------------------------------
    功能说明  : 段表驱动，一次调用把源 128 位窗口里的至多 8 个位段搬到目标窗口的指定
                位置（位段可跨 32 位字边界）。库内 BitArrayInsert 每次只能搬一段，
                多段场景要调用方自己循环并托管中间量，本件即补此缺口；
                核心防御是「先快照后写」：先把所有段值读进快照数组，全部读完后统一
                写目标，杜绝「段 1 的写覆盖段 2 的源」这类顺序缺陷；
                第二道防御是「逐位搬运」，任何宽度都不需要 32 位整字移位，
                彻底规避移位量等于 32 的未定义行为；
                越界段绝不部分写入，只跳过并计数；目标段重叠按段序后者覆盖前者并提示。
    错误码    : 16#0001_023B 存在越界 / 重叠段，已跳过并计数——信息级，正常防御
                16#0001_023C 预留禁用（信息级，不得挪用）
                16#0001_030F 段数为 0 或宽度全为 0——故障级，本拍不搬运
                16#0001_0310 段表自相矛盾（段数超段表容量）——故障级，本拍不搬运
                16#0001_0311 循环守卫超限（防死锁计数触发）——故障级，本拍结果作废
    码位总账  : 16#0001_023B 用 / 16#0001_023C 预留 ｜ 16#0001_030F 用 / 16#0001_0310 用 / 16#0001_0311 用
    状态机    : N/A —— 纯函数无顺序状态机，无 CASE 可写，非法状态不可能出现
    采样约定  : 纯组合函数，无定时器、无内部驻留状态，调用即出结果；
                目标窗口由调用方通过 VAR_IN_OUT 注入，本件绝不初始化目标数组。
    修订记录  : 2026-11-16 v1.0.0 首次入库（R18）
*)
FUNCTION FC_DL_BitSegmentBlockMove : BOOL
VAR_INPUT
    auSrcBit  : ARRAY[0..7] OF UINT;           // 各段源起始位（相对 128 位窗口）[位]，范围 0~127 / segment source start bit in the 128-bit window [bit], range 0~127
    auDstBit  : ARRAY[0..7] OF UINT;           // 各段目标起始位 [位]，范围 0~127 / segment destination start bit [bit], range 0~127
    auWidth   : ARRAY[0..7] OF UINT;           // 各段宽度 [位]，范围 1~32 / segment width [bit], range 1~32
    uSegCount : UINT := 1;                     // 有效段数 [段]，范围 1~8 / valid segment count [seg], range 1~8
    auSrcWord : ARRAY[0..3] OF DWORD;          // 源 128 位窗口，索引 0 = 最低字 [位图] / source 128-bit window, index 0 = lowest word [bitmap]
END_VAR
VAR_IN_OUT
    auDstWord : ARRAY[0..3] OF DWORD;          // 目标 128 位窗口，由调用方注入，本件不初始化 [位图] / destination window injected by the caller, never initialised here [bitmap]
END_VAR
VAR_OUTPUT
    uMovedSeg   : UINT;                        // 实际搬运段数 [段] / segments actually moved [seg]
    uSkippedSeg : UINT;                        // 因越界 / 重叠被跳过的段数 [段] / segments skipped due to range or overlap [seg]
    eErr        : UDINT;                       // 错误码，0=正常 / error id, 0=ok
    bError      : BOOL;                        // 故障标志，eErr 为故障级时 TRUE / error flag, TRUE on fault-level eErr
END_VAR
VAR
    uSeg      : UINT;                          // 段游标 [段] / segment cursor [seg]
    uBit      : UINT;                          // 段内位游标 [位] / bit cursor inside a segment [bit]
    uWr       : UINT;                          // 已写段遍历游标 [段] / written segment traversal cursor [seg]
    uGuard    : UINT;                          // 循环守卫计数 [次] / loop guard counter [times]
    uSrcAbs   : UINT;                          // 源窗口绝对位号 [位] / absolute bit number in the source window [bit]
    uDstAbs   : UINT;                          // 目标窗口绝对位号 [位] / absolute bit number in the destination window [bit]
    uWordIdx  : UINT;                          // 字索引 0~3 [字] / word index 0~3 [word]
    uBitPos   : UINT;                          // 字内位号 0~31 [位] / bit position inside a word 0~31 [bit]
    uBitMask  : DWORD;                         // 单比特掩码 [位图] / single bit mask [bitmap]
    abUse     : ARRAY[0..7] OF BOOL;           // 段可用标志（宽度合法且判界通过）/ usable segment flag, width legal and range checked
    auSnap    : ARRAY[0..7] OF DWORD;          // 段值快照，先快照后写 [位图] / segment value snapshot, read all before writing any [bitmap]
    auWrStart : ARRAY[0..7] OF UINT;           // 已写段起始位，重叠检测用 [位] / written segment start bit for overlap detection [bit]
    auWrEnd   : ARRAY[0..7] OF UINT;           // 已写段结束位，重叠检测用 [位] / written segment end bit for overlap detection [bit]
    uWrCnt    : UINT;                          // 已写段计数 [段] / written segment count [seg]
    bOverlap  : BOOL;                          // 本段与已写段重叠标志 / overlap flag against the written segments
    uValidN   : UINT;                          // 宽度合法的段数 [段] / segments with a legal width [seg]
END_VAR
VAR CONSTANT
    DL_SEG_MAX      : UINT := 8;               // 段表容量上限 [段] / segment table capacity [seg]
    DL_SEG_WIN_BITS : UINT := 128;             // 窗口位宽 [位] / window width [bit]
    DL_SEG_WORD_BITS: UINT := 32;              // 单字位宽 [位] / word width [bit]
    DL_SEG_MAX_LOOP : UINT := 8;               // 循环守卫硬上限 [次] / hard loop guard limit [times]
    DL_SEG_WIDTH_MAX: UINT := 32;              // 单段最大宽度 [位] / maximum single segment width [bit]
    DL_SEG_BIT_ONE  : DWORD := 16#0000_0001;   // 最低位掩码，移位量恒小于 32 [位图] / least significant bit mask, shift count always below 32 [bitmap]
END_VAR

// 段 1｜返回值与错误状态预置 / segment 1, preset return value and error status
FC_DL_BitSegmentBlockMove := FALSE;            // 故障缺省返回 FALSE / fault default returns FALSE
eErr := 0;                                     // 预置无错误 / preset no error
bError := FALSE;                               // 预置无故障 / preset no fault
uMovedSeg := 0;                                // 搬运段数清零 / clear the moved count
uSkippedSeg := 0;                              // 跳过段数清零 / clear the skipped count
uWrCnt := 0;                                   // 已写段计数清零 / clear the written count
uValidN := 0;                                  // 合法宽度段数清零 / clear the legal width count
uGuard := 0;                                   // 守卫计数清零 / clear the guard counter

// 段 2｜段数闸：0 段与超容量分别归入两个故障码，绝不索引越界 / segment 2, segment count gate
IF uSegCount < 1 THEN
    eErr := 16#0001_030F;                      // 段数为 0 故障码 / zero segment count fault id
    bError := TRUE;                            // 置故障标志 / raise the error flag
    RETURN;                                    // 故障级提前返回 / early return on fault
END_IF
IF uSegCount > DL_SEG_MAX THEN
    eErr := 16#0001_0310;                      // 段表自相矛盾故障码 / contradictory segment table fault id
    bError := TRUE;                            // 置故障标志 / raise the error flag
    RETURN;                                    // 故障级提前返回 / early return on fault
END_IF

// 段 3｜段表预清与宽度预筛：宽度不在 1~32 的段直接判不可用 / segment 3, clear the table and pre-screen the widths
FOR uSeg := 0 TO DL_SEG_MAX - 1 DO
    abUse[uSeg] := FALSE;                      // 先全部判不可用 / mark every segment unusable first
    auSnap[uSeg] := 0;                         // 快照清零 / clear the snapshot
    auWrStart[uSeg] := 0;                      // 写区间记录清零 / clear the written range start
    auWrEnd[uSeg] := 0;                        // 写区间记录清零 / clear the written range end
END_FOR
FOR uSeg := 0 TO uSegCount - 1 DO
    IF (auWidth[uSeg] >= 1) AND (auWidth[uSeg] <= DL_SEG_WIDTH_MAX) THEN
        abUse[uSeg] := TRUE;                   // 宽度合法，进入判界 / legal width, proceed to the range check
        uValidN := uValidN + 1;                // 合法段计数 / count the legal segment
    END_IF
END_FOR
IF uValidN < 1 THEN
    eErr := 16#0001_030F;                      // 宽度全为 0 故障码 / all widths zero fault id
    bError := TRUE;                            // 置故障标志 / raise the error flag
    RETURN;                                    // 故障级提前返回 / early return on fault
END_IF

// 段 4｜第一遍：判界 + 快照读（此遍绝不写目标）/ segment 4, first pass, range check and snapshot read only
FOR uSeg := 0 TO uSegCount - 1 DO
    uGuard := uGuard + 1;                      // 守卫累加 / accumulate the guard
    IF uGuard > DL_SEG_MAX_LOOP THEN
        eErr := 16#0001_0311;                  // 守卫超限故障码 / guard exceeded fault id
        bError := TRUE;                        // 置故障标志 / raise the error flag
        RETURN;                                // 结果作废 / discard the whole result
    END_IF
    IF abUse[uSeg] THEN
        IF ((auSrcBit[uSeg] + auWidth[uSeg]) > DL_SEG_WIN_BITS)
           OR ((auDstBit[uSeg] + auWidth[uSeg]) > DL_SEG_WIN_BITS)
           OR (auSrcBit[uSeg] >= DL_SEG_WIN_BITS)
           OR (auDstBit[uSeg] >= DL_SEG_WIN_BITS) THEN
            abUse[uSeg] := FALSE;              // 越界段判不可用，绝不部分写入 / out-of-range segment unusable, never partially written
            uSkippedSeg := uSkippedSeg + 1;    // 跳过计数 / count the skip
            eErr := 16#0001_023B;              // 越界提示（信息级不置故障）/ range hint, info level never raises a fault
        ELSE
            FOR uBit := 0 TO auWidth[uSeg] - 1 DO
                uSrcAbs := auSrcBit[uSeg] + uBit;             // 源绝对位号 / absolute source bit
                uWordIdx := uSrcAbs / DL_SEG_WORD_BITS;        // 字索引，绝对位号不超过 127 故不超过 3 / word index, absolute bit never exceeds 127 so never exceeds 3
                uBitPos := uSrcAbs - uWordIdx * DL_SEG_WORD_BITS; // 字内位号 0~31 / bit position inside the word 0~31
                uBitMask := SHL(DL_SEG_BIT_ONE, uBitPos);      // 掩码，移位量恒小于 32 / mask, shift count always below 32
                IF (auSrcWord[uWordIdx] AND uBitMask) <> 0 THEN
                    auSnap[uSeg] := auSnap[uSeg] OR SHL(DL_SEG_BIT_ONE, uBit); // 位收敛进快照 / gather the bit into the snapshot
                END_IF
            END_FOR
        END_IF
    ELSE
        uSkippedSeg := uSkippedSeg + 1;        // 宽度非法段同样计数跳过 / count the illegal width segment as skipped
        eErr := 16#0001_023B;                  // 跳过提示（信息级不置故障）/ skip hint, info level never raises a fault
    END_IF
END_FOR

// 段 5｜第二遍：统一写目标（快照已完整，读写互不污染）/ segment 5, second pass, single write phase
FOR uSeg := 0 TO uSegCount - 1 DO
    IF abUse[uSeg] THEN
        bOverlap := FALSE;                     // 重叠标志先清 / clear the overlap flag
        FOR uWr := 0 TO uWrCnt - 1 DO
            IF (auDstBit[uSeg] < auWrEnd[uWr]) AND ((auDstBit[uSeg] + auWidth[uSeg]) > auWrStart[uWr]) THEN
                bOverlap := TRUE;              // 与已写区间相交 / overlaps a written range
            END_IF
        END_FOR
        IF bOverlap THEN
            eErr := 16#0001_023B;              // 重叠提示，按段序后者覆盖前者（信息级）/ overlap hint, later segment overwrites the earlier one (info level)
        END_IF
        FOR uBit := 0 TO auWidth[uSeg] - 1 DO
            uDstAbs := auDstBit[uSeg] + uBit;                  // 目标绝对位号 / absolute destination bit
            uWordIdx := uDstAbs / DL_SEG_WORD_BITS;            // 字索引，判界已保证不超过 3 / word index, guaranteed below 4 by the range check
            uBitPos := uDstAbs - uWordIdx * DL_SEG_WORD_BITS;  // 字内位号 0~31 / bit position inside the word 0~31
            uBitMask := SHL(DL_SEG_BIT_ONE, uBitPos);          // 掩码，移位量恒小于 32 / mask, shift count always below 32
            IF (auSnap[uSeg] AND SHL(DL_SEG_BIT_ONE, uBit)) <> 0 THEN
                auDstWord[uWordIdx] := auDstWord[uWordIdx] OR uBitMask;      // 置位 / set the bit
            ELSE
                auDstWord[uWordIdx] := auDstWord[uWordIdx] AND NOT uBitMask; // 清位 / clear the bit
            END_IF
        END_FOR
        auWrStart[uWrCnt] := auDstBit[uSeg];   // 记录本次写区间起点 / record the written range start
        auWrEnd[uWrCnt] := auDstBit[uSeg] + auWidth[uSeg]; // 记录本次写区间终点 / record the written range end
        uWrCnt := uWrCnt + 1;                  // 已写段加一，上界由段数闸保证 / increment the written count, bounded by the segment gate
        uMovedSeg := uMovedSeg + 1;            // 搬运段数加一 / increment the moved count
        uGuard := uGuard + 1;                  // 守卫累加 / accumulate the guard
        IF uGuard > (DL_SEG_MAX_LOOP * 2) THEN
            eErr := 16#0001_0311;              // 守卫超限故障码 / guard exceeded fault id
            bError := TRUE;                    // 置故障标志 / raise the error flag
            RETURN;                            // 结果作废 / discard the whole result
        END_IF
    END_IF
END_FOR

// 段 6｜出口：至少搬成一段且无故障级码才返回 TRUE / segment 6, exit with TRUE only when something moved and no fault occurred
FC_DL_BitSegmentBlockMove := (NOT bError) AND (uMovedSeg > 0); // 成败判据 / success criterion
END_FUNCTION

(* ---- FC_DL_BitSet.st ---- *)
(*==============================================================================
 * 组件名称 (Component)  : FC_DL_BitSet
 * 所属子库 (Sublibrary) : DL_Base
 * 当前版本 (Version)    : 1.0.0
 * 兼容性   (Platform)   : CODESYS 3.5 / TwinCAT 3 / 汇川 InoProShop / Machine Expert
 *                         仅用标准 SHL / AND / OR / NOT，无任何厂商位写语法
 * 功能描述 (Function)   : 对 32 位字做"置位 / 清零"的纯函数操作：输入原值、返回新值，
 *                         不修改入参、不产生副作用，可安全用于表达式与 CASE 分支链式调用。
 *                         位索引越界时"原样返回原字"（不做任何修改），并给出错误码——
 *                         返回 0 会把整个状态字清零，在报警字场景等同于"全部报警消失"，
 *                         属危险的静默失败。
 * 开源溯源 (Origin)     : 原创实现。掩码构造方式参照 IEC 61131-3 位串运算语义，
 *                         不使用任何 CODESYS / TwinCAT 专有位访问扩展。
 * 依赖     (Depends)    : 无 DL_ 内部依赖；无标准库功能块依赖
 * 红线自检 (Redline)    : R1 ✓ 零全局变量表与外部变量引用 ｜ R2 ✓ 零物理 IO 地址直写
 *                         R3 ✓ 纯 IEC 61131-3（无厂商位写方言）｜ R4 ✓ 越界原样返回 + 掩码后构造
 *                         R5 ✓ 全变量中英双语同行注释 ｜ R6 N/A（无状态机）｜ R7 N/A（无实例调用）
 * 修订历史 (Revision)   :
 *   2026-11-14  v1.0.0  首版入库（Phase 1 冷启动 · Level 0 批次）
 *============================================================================*)
FUNCTION FC_DL_BitSet : DWORD
VAR_INPUT
    uValue    : DWORD;             // 原始状态字，函数内只读 / Source status word, read-only inside the function
    uBitIndex : USINT;             // 位序号，0 = LSB，合法域 0..31 / Bit index, 0 = LSB, valid range 0..31
    bSetValue : BOOL := TRUE;      // TRUE = 置 1，FALSE = 清 0 / TRUE = set to 1, FALSE = clear to 0
END_VAR
VAR_OUTPUT
    bValid    : BOOL;              // 索引合法标志，FALSE 时返回原值 / Index valid flag, FALSE means the input is returned unchanged
    uErrorId  : UDINT;             // 故障码，0 = 无故障 / Error code, 0 = no error
END_VAR
VAR
    uMask      : DWORD;            // 目标单位掩码 / Single-bit target mask
    uWorkValue : UDINT;            // 提升到 UDINT 的原值工作副本 / UDINT working copy of the source value
    uWorkMask  : UDINT;            // 提升到 UDINT 的掩码工作副本 / UDINT working copy of the mask
    uShift     : UDINT;            // 提升到 UDINT 的移位量 / Shift amount promoted to UDINT
END_VAR
VAR CONSTANT
    DL_BIT_INDEX_MAX : USINT := 31;  // 32 位字的最大合法位索引 / Max legal bit index of a 32-bit word
END_VAR

(*------------------------------------------------------------------------------
 * 段 1｜返回值预置为原值（边界 B1）：异常路径下"不做任何修改"是最安全语义
 *      Pre-set return to the source value: on any error path, "change nothing" is safest
 *-----------------------------------------------------------------------------*)
FC_DL_BitSet := uValue;
bValid       := FALSE;
uErrorId     := 16#0000_0000;
uMask        := 16#0000_0000;
uWorkValue   := 16#0000_0000;
uWorkMask    := 16#0000_0000;
uShift       := 16#0000_0000;

(*------------------------------------------------------------------------------
 * 段 2｜越界拦截：先校验、后构造掩码（边界 B2，顺序即防御）
 *      Bounds interception: validate first, build the mask afterwards
 *      越界时立即返回原值，绝不执行 SHL(1, index) 以免触发未定义行为
 *-----------------------------------------------------------------------------*)
IF uBitIndex > DL_BIT_INDEX_MAX THEN
    uErrorId := 16#0001_0001;
    RETURN;
END_IF

(*------------------------------------------------------------------------------
 * 段 3｜掩码构造：UDINT#1 左移 index 位，得到仅目标位为 1 的单位掩码
 *      Mask construction: shift UDINT#1 by index to obtain a single-bit mask
 *      使用显式类型字面量 UDINT#1，避免隐式类型转换（红线 R3）
 *-----------------------------------------------------------------------------*)
uShift    := USINT_TO_UDINT(uBitIndex);
uWorkMask := SHL(UDINT#1, uShift);
uMask     := UDINT_TO_DWORD(uWorkMask);
uWorkValue := DWORD_TO_UDINT(uValue);

(*------------------------------------------------------------------------------
 * 段 4｜置位 / 清零（边界 B3）：两条路径共用同一掩码，保证完全对称
 *      Set / clear: both paths share one mask, guaranteeing symmetry
 *      清零用 AND NOT 作用于 UDINT 全域 32 位，不得只反低 8 位而误伤其它位
 *-----------------------------------------------------------------------------*)
IF bSetValue THEN
    uWorkValue := uWorkValue OR uWorkMask;
ELSE
    uWorkValue := uWorkValue AND NOT uWorkMask;
END_IF

(*------------------------------------------------------------------------------
 * 段 5｜结果回写：经返回值输出，入参 uValue 全程未被修改（边界 B4）
 *      Result write-back through the return value, the input stays untouched
 *-----------------------------------------------------------------------------*)
FC_DL_BitSet := UDINT_TO_DWORD(uWorkValue);
bValid       := TRUE;
END_FUNCTION

(* ---- FC_DL_BitSwapPairs.st ---- *)
(*==============================================================================
 * 名称 : FC_DL_BitSwapPairs —— BYTE 内相邻比特对交换（4 对：0↔1,2↔3,4↔5,6↔7）
 * 分类 / 前缀 / 版本 : DL_Base / FC_DL_ / 1.0.0
 * 溯源 : 开源语义参考（OSCAT/AixOCAT 族，MIT）或 clean-room IEC 实现，未复制源码
 * 平台 : 纯 IEC 61131-3
 * 功能说明 : 将 BYTE 的 4 个相邻位对两两交换后返回：偶数位整体左移 1、奇数位
 *            整体右移 1，再按位或合成（掩码 16#55 取偶位、16#AA 取奇位）。
 *            边界处理：全 0 / 全 1 / 对称位型（如 16#66）交换后为原值，属合法
 *            结果；移位量恒 1（< 8 位宽），结构性无越界移位。
 * 错误码 : 无故障路径（全值域合法的纯变换），eErr 恒 0，bValid 恒 TRUE；
 *          16#0001_1A06 为本件预留码位，当前实现不发出
 * 状态机 : R6 标注 N/A（纯函数无顺序状态，以本节替代 ELSE 兜底）
 * 红线 : R1/R2/R3 ✓ 零全局/零IO/纯IEC ｜ R4 ✓ 移位量=1 ｜ R10 ✓ 标准转换 ｜ R11 ✓ 分号收尾 ｜ R15 ✓ 无保留字撞名
 * 修订记录 : 2026-11-23 v1.0.0 首次入库（R76）
 *============================================================================*)
FUNCTION FC_DL_BitSwapPairs : BYTE
VAR_INPUT
    byIn : BYTE;       // 待交换的输入字节 [位域] / input byte for pair swap
END_VAR
VAR_OUTPUT
    eErr   : UDINT;    // 故障码，0=正常（本件无故障路径）/ error code, 0=ok (no fault path)
    bError : BOOL;     // 故障标志，恒 FALSE / error flag, always FALSE
    bValid : BOOL;     // TRUE=返回值可用，恒 TRUE / TRUE when return value is usable
END_VAR
VAR
    _byEven : BYTE;    // 偶数位左移后的分量 [位域] / even-bit component shifted left
    _byOdd  : BYTE;    // 奇数位右移后的分量 [位域] / odd-bit component shifted right
END_VAR

eErr   := 16#0000_0000;                      // 故障码清零 / clear error code
bError := FALSE;                             // 故障标志清零 / clear error flag
bValid := TRUE;                              // 本件全值域合法，恒可用 / always valid

_byEven := SHL(byIn AND BYTE#16#55, 1);      // 偶位掩码后左移 1 位（<8 安全）/ even bits shifted up by one
_byOdd  := SHR(byIn AND BYTE#16#AA, 1);      // 奇位掩码后右移 1 位（<8 安全）/ odd bits shifted down by one
FC_DL_BitSwapPairs := _byEven OR _byOdd;     // 两分量按位或合成 / compose by bitwise or

END_FUNCTION

(* ---- FC_DL_ByteArrayXor.st ---- *)
(*==============================================================================
 * 组件名称 (Component)  : FC_DL_ByteArrayXor
 * 所属子库 (Sublibrary) : DL_Base
 * 当前版本 (Version)    : 1.0.0
 * 兼容性   (Platform)   : CODESYS 3.5+ / TwinCAT 3 / 汇川 InoProShop / 施耐德 Machine Expert
 *                         仅依赖 IEC 61131-3 位运算内建，零厂商私有库
 * 功能描述 (Function)   : 字节数组异或校验和（BCC / Block Check Character），用于串口协议帧尾校验。
 *                         逐字节按序异或，结果 BYTE 单字节出口。
 *                         与 CRC16-Modbus / LRC 件的差别（属主边界）：BCC 是无进位单字节异或，
 *                         无初值/无反射/无多项式，不可互替；三者各占一件，判据互不共用。
 *                         验收向量（算法级自证，脚本可复算）：
 *                           ① 空数组 uLen=0            → 拒算返回 16#00 + bInvalid
 *                           ② {16#55}                  → 16#55
 *                           ③ {16#01, 16#02, 16#03}    → 16#00（1^2=3，3^3=0，异或自反性）
 *                           ④ {16#FF, 16#F0}           → 16#0F
 * 接口     (Interface)  : 入 aBytes 待校验字节缓冲（IN_OUT，调用者持有）、uLen 有效长度；
 *                         出 返回值 = BCC 字节、bInvalid 拒算标志、bClamped 长度越上限钳位标志。
 * 边界     (Boundary)   : ① **空数组拒算**：uLen = 0 → 返回 16#00 + bInvalid（空帧的异或和为 0
 *                         会与"单字节 0"不可区分，是伪校验，故拒算而非返回真值）；
 *                         ② **长度上限防扫爆**：uLen > 256 时钳到 256 并置 bClamped，
 *                         不允许调用者声明的长度把循环拖进长扫描（R104 运行时二次闸）；
 *                         ③ 数组上界以**字面量 255** 声明（接口上界须编译期常量，R104），
 *                         同值常量 DL_BCC_MAX_LEN=256 作运行时二次闸，两处同源、改动须同步；
 *                         ④ 调用者须保证 uLen ≤ 实际数组长度（IN_OUT 语义，本件只做上限侧防御）；
 *                         ⑤ 纯函数无记忆量；零全局耦合、零物理地址。
 * 分工声明 (Scope)      : 本件只管"单字节异或和"。不接管：CRC/LRC 多项式校验、帧头帧长解析、
 *                         校验失败后的重发编排（属协议层件）。
 * 来源标签 (Source Tag) : T0 防御包装 —— IEC 61131-3 标准语义的道莅防御性实现
 * 码表     (Codes)      : 本件不占用任何全局数字码位（零码位范式 R297）；诊断由 BOOL 出口承担。
 * 红线自检 (Redline)    : R1 ✓ 零 GVL/VAR_EXTERNAL ｜ R2 ✓ 零 %I/%Q/%M ｜ R3 ✓ 纯 IEC 61131-3
 *                         R4 ✓ 空数组闸 + 长度上限钳 + 双端循环上界 ｜ R5 ✓ 声明逐行同行双语注释
 *                         R6 ✓ 无状态机（纯组合函数，判别用 IF 链含两分支） ｜ R7 ✓ 无定时器/沿实例
 * 修订历史 (Revision)   : 2026-11-19  v1.0.0  R47 首版（批次 1 · 序号 2）
 *==============================================================================*)

FUNCTION FC_DL_ByteArrayXor : BYTE
VAR_IN_OUT
    aBytes : ARRAY[0..255] OF BYTE;         // 待校验字节缓冲（上界字面量，R104） [-] / Source byte buffer, literal bound
END_VAR
VAR_INPUT
    uLen : UINT := 0;                       // 有效字节数，域 0..256（0 拒算） [-] / Valid byte count, 0 rejected
END_VAR
VAR_OUTPUT
    bInvalid : BOOL := FALSE;               // 拒算标志（uLen=0，当拍有效） [-] / Rejection flag (uLen=0, this scan)
    bClamped : BOOL := FALSE;               // 长度越上限钳位标志 [-] / Length clamp flag (upper bound hit)
END_VAR
VAR
    uXor    : BYTE := 16#00;                // 异或累加器（初值 0 为异或单位元） [-] / XOR accumulator
    uLenUse : UINT := 0;                    // 归一后的实际扫描长度 [-] / Normalised scan length
    i       : UINT := 0;                    // 字节下标 / Byte index
END_VAR
VAR CONSTANT
    DL_BCC_MAX_LEN : UINT := 256;           // 扫描长度上限（与接口字面量上界 255 同源） [-] / Max scan length
END_VAR

(* —— 段 1：返回值与两标志预置（R45 四段式第①段） —— *)
FC_DL_ByteArrayXor := 16#00;                // 返回值预置异或单位元 / Return value preset to XOR identity
bInvalid := FALSE;                          // 拒算标志预置 / Rejection flag preset
bClamped := FALSE;                          // 钳位标志预置 / Clamp flag preset
uXor    := 16#00;                           // 累加器预置 / Accumulator preset
uLenUse := 0;                               // 长度工作量预置 / Length working value preset

(* —— 段 2：域闸门早退（空数组不扫、不宣称校验和） —— *)
IF uLen = 0 THEN
    bInvalid := TRUE;                       // 空数组拒算 / Empty array rejected
    FC_DL_ByteArrayXor := 16#00;            // 拒算返回值 / Return value on rejection
    RETURN;                                 // 早退，不进入扫描 / Early return, no scan
END_IF

(* —— 段 3：长度上限钳位（运行时二次闸，防调用者传巨值扫爆） —— *)
uLenUse := uLen;                            // 取调用者长度 / Take the caller length
IF uLenUse > DL_BCC_MAX_LEN THEN
    uLenUse := DL_BCC_MAX_LEN;              // 钳到上限 / Clamp to the upper bound
    bClamped := TRUE;                       // 置钳位标志 / Raise the clamp flag
END_IF

(* —— 段 4：逐字节异或（双端上界：uLenUse ≤ 256，下标恒在数组域内） —— *)
i := 0;                                     // 下标归零 / Index reset
WHILE (i < uLenUse) AND (i < DL_BCC_MAX_LEN) DO
    uXor := uXor XOR aBytes[i];             // 累加异或 / Accumulate XOR
    i := i + 1;                             // 计数器推进（循环必然收敛） / Counter advance, loop terminates
END_WHILE

(* —— 段 5：统一出口（BYTE 域天然闭合，无需再钳） —— *)
FC_DL_ByteArrayXor := uXor;                 // 输出 BCC 单字节 / Output the BCC byte

END_FUNCTION

(* ---- FC_DL_BytesToWord.st ---- *)
(*==============================================================================
 * 名称 : FC_DL_BytesToWord —— 双字节按序组装 WORD（显式大小端参数）
 * 分类 / 前缀 / 版本 : DL_Base / FC_DL_ / 1.0.0
 * 溯源 : 开源语义参考（OSCAT/AixOCAT 族，MIT）或 clean-room IEC 实现，未复制源码
 * 平台 : 纯 IEC 61131-3
 * 功能说明 : 将高/低两个 BYTE 按 bBigEndian 指定的顺序组装为 WORD：大端时
 *            byHi 为高 8 位、byLo 为低 8 位；小端时两者角色对调。
 *            装配全程使用数值语义（BYTE_TO_WORD + SHL/AND/OR），不触碰内存序。
 *            边界处理：byHi/byLo 全值域合法（BYTE 天然 ≤255），无溢出可能。
 * 错误码 : 无故障路径（全值域合法的纯装配），eErr 恒 0，bValid 恒 TRUE；
 *          16#0001_1A09 为本件预留码位，当前实现不发出
 * 状态机 : R6 标注 N/A（纯函数无顺序状态，以本节替代 ELSE 兜底）
 * 红线 : R1/R2/R3 ✓ 零全局/零IO/纯IEC（禁指针/联合体）｜ R4 ✓ 移位量=8 ｜ R10 ✓ 标准转换 ｜ R11 ✓ 分号收尾 ｜ R15 ✓ 无保留字撞名
 * 修订记录 : 2026-11-23 v1.0.0 首次入库（R76）
 *============================================================================*)
FUNCTION FC_DL_BytesToWord : WORD
VAR_INPUT
    byHi       : BYTE;     // 语义高位字节 [0..255] / semantically high byte
    byLo       : BYTE;     // 语义低位字节 [0..255] / semantically low byte
    bBigEndian : BOOL;     // TRUE=大端装配（byHi 在高位）/ TRUE for big-endian assembly
END_VAR
VAR_OUTPUT
    eErr   : UDINT;    // 故障码，0=正常（本件无故障路径）/ error code, 0=ok (no fault path)
    bError : BOOL;     // 故障标志，恒 FALSE / error flag, always FALSE
    bValid : BOOL;     // TRUE=返回值可用，恒 TRUE / TRUE when return value is usable
END_VAR
VAR
    _wH : WORD;        // 高字节拓宽值 [0..255] / widened high byte
    _wL : WORD;        // 低字节拓宽值 [0..255] / widened low byte
END_VAR

eErr   := 16#0000_0000;                      // 故障码清零 / clear error code
bError := FALSE;                             // 故障标志清零 / clear error flag
bValid := TRUE;                              // 本件全值域合法，恒可用 / always valid

_wH := BYTE_TO_WORD(byHi);                   // 高字节零拓宽至 16 位（无符号安全）/ widen high byte zero-extended
_wL := BYTE_TO_WORD(byLo);                   // 低字节零拓宽至 16 位（无符号安全）/ widen low byte zero-extended

IF bBigEndian THEN                           // 大端：byHi 占高 8 位 / big-endian: byHi goes high
    FC_DL_BytesToWord := SHL(_wH, 8) OR _wL; // 高字节左移 8 位后并入低字节（移位量 8<16 安全）/ compose
ELSE                                         // 小端：byLo 占高 8 位 / little-endian: byLo goes high
    FC_DL_BytesToWord := SHL(_wL, 8) OR _wH; // 低字节左移 8 位后并入高字节 / compose swapped
END_IF

END_FUNCTION

(* ---- FC_DL_DaysInMonthChk.st ---- *)
(*
    FC_DL_DaysInMonthChk —— 年月 → 当月天数（日历原子族补件）
    ------------------------------------------------------------------
    组件名称  : FC_DL_DaysInMonthChk
    分类      : DL_Base / Calendar
    前缀      : FC_DL_
    版本      : 1.0.0
    溯源      : IEC 61131-3 标准语义的道莅防御性实现（格里高利历月天数
                静态表 + 闰年二月分支）；闰年律**唯一属主为库内
                FC_DL_LeapYearChk（DL_Base），本件组合调用之，零内联
                4/100/400 三级判定（常量单源纪律）**；月天数表为公开历法
                常识；实现 / 引脚名 / 码位 100% 自有；clean-room 声明 ——
                零代码行复制，无闭源参考。
    平台      : 纯 IEC 61131-3（CASE + 组合调用），无内建函数依赖，
                CODESYS 3.5 / TwinCAT 3 / InoProShop / Machine Expert 通用
    作者      : 道莅代码库 · PLC编程专家（R72 构建轮 · 批 3 · 序号 7）
    ------------------------------------------------------------------
    功能说明  : 年月 → 当月天数（28~31 四值）。真实工况：月末日期计算、
                月度报表界、计量月切账日推演。
                判据链顺序：
                ① 年份承诺段闸：**[1998, 2099]**，域外故障级拒绝、输出 0、
                   不钳位照算——月天数是日历**事实**而非量值（R81 还原方向
                   不饱和：对域外年份伪造天数会一路传到月末日期运算）；
                ② 月域闸：1~12 外 → 故障级早退输出 0；
                ③ 大小月静态表出口（31 / 30）；
                ④ 二月分支：**组合调用闰年律唯一属主 FC_DL_LeapYearChk
                   （bFullRule := TRUE 三律，2000 世纪年判闰的事实正确性由
                   三律保证）**，属主件信息级 0430（整百年）在无更高优先级
                   码时透传；属主回执防御收口（不可达）。
                计划偏差声明（留痕）：ROUND_PLAN_R72 §6 承诺段写 1998~2117
                （DATE 容器秒承载口径），实测属主件闰年窗口为 1900~2099，
                本件承诺段**收窄对齐为 [1998, 2099]**；2100~2117 请求按 R81
                事实口径故障级拒绝而非钳位（钳位 2099 会把 2104 闰年误报为
                平年 28 天——钳位即伪造事实，故拒绝），偏差已留 VERSION 口径。
    错误码    : 16#0001_0750 月域越界（<1 或 >12），输出 0 —— 故障级
                16#0001_0751 年份越承诺段 [1998, 2099]，输出 0，不钳位
                            （R81 事实口径）—— 故障级
                16#0001_0753 闰年属主件回执不可用（年份已预闸入属主窗口，
                            结构性不可达防御收口）—— 故障级
                16#0001_0430（属主件信息级透传）整百年，闰年结论取决于三律
                            —— 信息级，不置 bError（R45）
                加码反证句（R90）：0750 / 0751 由入参域直接可证互斥观测；
                0753 与 0751 输出同为 0 + 故障级，但 0751 的入参越域可被
                调用方自证、0753 的入参合法，成因互斥不可互换，故各立一码。
    码位总账  : 16#0001_0750 用 ｜ 16#0001_0751 用 ｜ 16#0001_0753 用
                （16#0001_0752 为同段邻件 FB_DL_BlinkOutput 组态锁存码，
                本件不用不占）
    状态机    : N/A —— 纯函数无状态；月分支用 CASE + ELSE 兜底（月闸后
                ELSE 结构性不可达，防御收口并入 0750）
    边界与披露: 一 无定时器 / 无沿检测实例 / 无数组下标 / 无除法 / 无循环，
                   周期安全规则 N/A；
                二 零全局变量、零 VAR_EXTERNAL、零物理地址；
                三 整数进位点（终审两式 #2）验收向量：月域「1 恰为下界」
                   → 31 合法出口；「0 / 13 越界」→ 0750 故障级；闰年向量
                   三组（2024 闰 → 29 / 2100 世纪非闰 → 0751 拒绝出域 /
                   2000 闰 → 29 + 0430 透传）随验收落 JSONL；
                四 域闸逐项点名（R272）：uYear / uMonth 两入参全部纳入域闸；
                五 归位声明：日历 FC 原子族（LeapYearChk / DayOfWeekCalc /
                   WeekOfYearCalc / DurationFormat）属主均在 DL_Base
                   （registry 实测），本件随族归位；
                六 分工互引：FC_DL_LeapYearChk（闰年律唯一属主）、
                   FB_DL_MonthWindowCheck（月窗判定，可消费本件简化月末界）
                   ——本件只做月天数原子；
                七 依赖声明：仅 Standard.library（无内建函数依赖）+ 同库
                   FC_DL_LeapYearChk（只调用不修改）。
    验收向量  : V1 (2024, 2) → 29；V2 (2100, 2) → 0751 故障级输出 0；
                V3 (2000, 2) → 29 + 0430 信息级透传；V4 (2023, 4) → 30；
                V5 (2023, 7) → 31；V6 (2020, 1) → 31（年合法月下界 1 恰过闸）；
                V7 (2020, 0) / (2020, 13) → 0750 故障级输出 0；
                V8 (1997, 2) / (2099, 2) → 承诺段两端点（1997 拒 0751，
                2099 平年 → 28）。
                算法已证（脚本）：未跑 ｜ 编译器已证（三平台）：未跑
    修订记录  : 2026-11-23 v1.0.0 首次入库（R72 构建轮 · 批 3 · 序号 7）
*)
FUNCTION FC_DL_DaysInMonthChk : USINT
VAR_INPUT
    uYear  : UINT;                         (* 年份，[年]，承诺段 [1998, 2099]（与闰年属主窗口对齐收窄），域外拒绝不钳位 / the year, promise range 1998 to 2099, refused outside *)
    uMonth : UINT;                         (* 月份，[月]，域 [1, 12]，域外拒绝 / the month, domain 1 to 12, refused outside *)
END_VAR
VAR_OUTPUT
    bValid    : BOOL;                      (* 返回值（天数）可用标志，故障级为 FALSE / the days usable flag *)
    bError    : BOOL;                      (* 故障标志，仅故障级码置位（R45 配对）/ the fault flag *)
    nInfoCode : UDINT;                     (* 信息 / 错误码，0 = 正常 / the info or error id *)
END_VAR
VAR CONSTANT
    DL_DIM_YMIN  : UINT := 1998;           (* 年份承诺段下界 [年] / the year promise lower bound *)
    DL_DIM_YMAX  : UINT := 2099;           (* 年份承诺段上界（属主闰年窗口对齐收窄）[年] / the year promise upper bound, aligned with the owner window *)
    DL_DIM_MMIN  : UINT := 1;              (* 月域下界 [月] / the month domain lower bound *)
    DL_DIM_MMAX  : UINT := 12;             (* 月域上界 [月] / the month domain upper bound *)
    DL_DIM_FEB   : UINT := 2;              (* 二月月号（闰年分支入口）[月] / the February selector *)
    DL_DIM_DAYS31: USINT := 31;            (* 大月天数 [日] / the big month days *)
    DL_DIM_DAYS30: USINT := 30;            (* 小月天数 [日] / the small month days *)
    DL_DIM_DAYS29: USINT := 29;            (* 闰二月天数 [日] / the leap February days *)
    DL_DIM_DAYS28: USINT := 28;            (* 平二月天数 [日] / the common February days *)
END_VAR
VAR
    _bLpyOk   : BOOL;                      (* 闰年属主件返回值回执（TRUE = 闰年）[标志] / the leap year owner return receipt *)
    _bLpyErr  : BOOL;                      (* 闰年属主件故障回执 [标志] / the leap year owner fault receipt *)
    _bLpyVld  : BOOL;                      (* 闰年属主件判定有效回执（R381 全回执）[标志] / the leap year owner verdict valid receipt *)
    _eLpyCode : UDINT;                     (* 闰年属主件码位回执 [码] / the leap year owner code receipt *)
    uDays     : USINT;                     (* 月天数工作副本 [日] / the days working copy *)
END_VAR

// 段 1｜返回值与状态预置（统一出口预置，R256）/ segment 1, preset the return and the status
FC_DL_DaysInMonthChk := 0;                 // 故障缺省返回 0 天 / the fault default is zero days
bValid    := FALSE;                        // 预置不可用，过闸后置位 / preset unusable
bError    := FALSE;                        // 预置无故障 / preset no fault
nInfoCode := 0;                            // 预置无错 / preset no error
_bLpyOk := FALSE;                          // 属主回执清零 / clear the owner receipts
_bLpyErr := FALSE;                         // 属主回执清零 / clear the owner receipts
_bLpyVld := FALSE;                         // 属主回执清零 / clear the owner receipts
_eLpyCode := 0;                            // 属主码位清零 / clear the owner code
uDays := 0;                                // 天数副本清零 / clear the days copy

// 段 2｜年份承诺段闸：域外拒绝不钳位（R81 事实口径，防伪造天数）/ segment 2, the year promise gate, refusal over clamping
IF (uYear < DL_DIM_YMIN) OR (uYear > DL_DIM_YMAX) THEN // 年份越承诺段 / the year out of the promise
    nInfoCode := 16#0001_0751;             // 故障级：年份越承诺段 / fault level: the year out of promise
    bError := TRUE;                        // R45 配对置故障标志 / paired with the fault flag
    bValid := FALSE;                       // 返回值不可用 / unusable
    FC_DL_DaysInMonthChk := 0;             // 确定值零出口 / a deterministic zero outlet
    RETURN;                                // 结构早退 / structural exit
END_IF

// 段 3｜月域闸：1~12 外故障级早退 / segment 3, the month domain gate
IF (uMonth < DL_DIM_MMIN) OR (uMonth > DL_DIM_MMAX) THEN // 月越域 / the month out of domain
    nInfoCode := 16#0001_0750;             // 故障级：月域越界 / fault level: the month out of domain
    bError := TRUE;                        // R45 配对置故障标志 / paired with the fault flag
    bValid := FALSE;                       // 返回值不可用 / unusable
    FC_DL_DaysInMonthChk := 0;             // 确定值零出口 / a deterministic zero outlet
    RETURN;                                // 结构早退 / exit
END_IF

// 段 4｜大小月静态表 + 二月闰年分支（CASE + ELSE 兜底，月闸后 ELSE 不可达）/ segment 4, the month table and the February leap branch
CASE uMonth OF
    1, 3, 5, 7, 8, 10, 12:                 // 大月组 / the big months
        uDays := DL_DIM_DAYS31;            // 31 天 / thirty one days
    4, 6, 9, 11:                           // 小月组 / the small months
        uDays := DL_DIM_DAYS30;            // 30 天 / thirty days
    DL_DIM_FEB:                            // 二月：复用闰年律唯一属主 / February, the leap law owner call
        _bLpyOk := FC_DL_LeapYearChk(nYear := uYear,    // 年份已预闸入属主窗口 [1998, 2099] / the year pre gated inside the owner window
                                     bFullRule := TRUE, // 三律（2000 世纪年判闰事实正确性）/ the full three rule set
                                     eErr => _eLpyCode, // 码位回执 / the code receipt
                                     bError => _bLpyErr, // 故障回执 / the fault receipt
                                     bValid => _bLpyVld); // 判定有效回执（R381 全回执）/ the verdict valid receipt
        IF (NOT _bLpyOk) OR _bLpyErr OR (NOT _bLpyVld) THEN // 属主回执防御收口（结构性不可达）/ the owner receipt defensive guard
            nInfoCode := 16#0001_0753;     // 故障级：属主回执不可用 / fault level: the owner receipt unusable
            bError := TRUE;                // R45 配对 / paired with the flag
            bValid := FALSE;               // 返回值不可用 / unusable
            FC_DL_DaysInMonthChk := 0;     // 确定值零出口 / a deterministic zero outlet
            RETURN;                        // 结构早退 / exit
        END_IF
        IF _bLpyOk THEN                    // 属主判闰 / the owner verdicts a leap year
            uDays := DL_DIM_DAYS29;        // 29 天 / twenty nine days
        ELSE                               // 属主判平 / the owner verdicts a common year
            uDays := DL_DIM_DAYS28;        // 28 天 / twenty eight days
        END_IF
        IF (nInfoCode = 0) AND (_eLpyCode <> 0) AND (NOT _bLpyErr) THEN // 属主信息级透传（无更高优先级码时）/ the owner info pass through
            nInfoCode := _eLpyCode;        // 信息级透传（0430 整百年提示）/ the info pass through
        END_IF
    ELSE                                   // 月闸后不可达防御兜底（并入 0750 口径）/ the unreachable ELSE after the month gate
        uDays := 0;                        // 确定值零出口 / a deterministic zero outlet
        nInfoCode := 16#0001_0750;         // 并入月域故障级（R90 反证：不可达无独立观测需求）/ folded into the month fault
        bError := TRUE;                    // R45 配对 / paired with the flag
        bValid := FALSE;                   // 返回值不可用 / unusable
        FC_DL_DaysInMonthChk := 0;         // 确定值零出口 / a deterministic zero outlet
        RETURN;                            // 结构早退 / exit
END_CASE

// 段 5｜正常出口 / segment 5, the normal outlet
FC_DL_DaysInMonthChk := uDays;             // 发布月天数（28~31）/ publish the days
bValid := TRUE;                            // 结果可用 / the result usable
END_FUNCTION

(* ---- FC_DL_DurationFormat.st ---- *)
(*
    FC_DL_DurationFormat —— TIME 时长分解为 天/时/分/秒 四分量（HMI 显示用纯函数）
    ------------------------------------------------------------------
    组件名称  : FC_DL_DurationFormat
    分类      : DL_Base / TimeFormat
    前缀      : FC_DL_
    版本      : 1.0.0
    溯源      : 借鉴点 —— IEC 61131-3 TIME 类型语义（无符号毫秒容器），
                T0-2 族内补口（Date and Timer → DL_Base 分类事实，T0 = 1，
                允许区间 0~1）。
                本件只借**标准类型语义**，分解规格与码位口径为自有。
                clean-room 声明 —— 零代码行复制；仅用标准类型转换
                TIME_TO_DINT / DINT_TO_UDINT 与整除 / 取模运算符。
                许可证 —— 本件 MIT。
    平台      : 纯 IEC 61131-3，CODESYS 3.5 / TwinCAT 3 / InoProShop / Machine Expert 通用
    作者      : 道莅代码库 · PLC编程专家（R71 构建轮 · 批 1 · 序号 4）
    ------------------------------------------------------------------
    功能说明  : 将输入时长 tDur 一次性换算到毫秒整数，再整除分解为
                天 / 时 / 分 / 秒四分量（HMI 显示口径，秒以下毫秒余量舍弃，
                向下取整到秒）：
                uDays  = uMs / 86400000，余数级联
                uHours = 余 / 3600000，余数级联
                uMins  = 余 / 60000，余数级联
                uSecs  = 余 / 1000，毫秒余量 = bTruncated 判据。
                除法除子全为**常量** 86400000 / 3600000 / 60000 / 1000
                （VAR CONSTANT 声明），**无变量除零面**（R45 纪律：常量除子
                不设判零闸，头注释声明即为口径）。
                负 TIME 不可表示（TIME 无符号语义）：输入域闸按防御性复检
                落码 —— TIME_TO_DINT 结果 < 0 即拒绝（非法入参），四分量
                清零、返回 FALSE；标准平台负 TIME 本就不可构造，闸属防御
                兜底而非业务判据（声明口径）。
                uDays 上界声明：TIME 容器毫秒上限 2147483647 ms（DINT 域）
                ÷ 86400000 = 24 天余 63487 秒分量 —— 四分量均为 UDINT，
                分解结果恒在容器内，无溢出面（声明即口径）。
    错误码    : N/A —— 本件按计划规格不出码位（输出契约：四分量 + bValid +
                bTruncated）；入参非法以返回值 FALSE 表达，四分量清零，
                绝不送未定义值给下游。
    码位总账  : 无码位（计划口径：多出口分解件，有效性以 bValid / 返回值承载）
    状态机    : N/A —— 纯函数无状态，无 CASE 可写，非法状态不可能出现
    边界与披露: 一 无定时器 / 无边沿实例 / 无数组下标，周期安全规则 N/A；
                二 零全局变量、零 VAR_EXTERNAL、零物理地址；
                三 整除分解全链无浮点量、无浮点判等面（纯整数运算）；
                四 bTruncated 语义：毫秒余量非零被舍弃（显示口径为向下取整
                   到秒），非「容器上界截断」—— TIME 入参本身即为容器
                   全域，不存在入参超出容器的问题（R191 名实双出口：
                   位名 bTruncated 对齐「余量舍弃」实现语义）；
                五 返回值即 bValid 语义（出参契约：入参合法且已完整分解
                   才 TRUE）。
    分工声明  : FC_DL_TimeToDintMs（DL_MathData，TIME → DINT 毫秒单一数值
                换算）、FC_DL_TimeToLrealSec（DL_MathData，TIME → LREAL 秒
                单一数值换算）—— 两者为**单一数值换算**件；本件为**日历
                分量分解**件（天 / 时 / 分 / 秒多出口语义，HMI 显示用），
                分工边界为「一个数 vs 四个分量」，非同算法变体，互引不互代。
    修订记录  : 2026-11-22 v1.0.0 首次入库（R71 构建轮 · 批 1 · 序号 4）
*)
FUNCTION FC_DL_DurationFormat : BOOL
VAR_INPUT
    tDur : TIME;                           (* 输入时长（TIME 无符号毫秒容器），[ms] / the input duration, an unsigned millisecond TIME container *)
END_VAR
VAR_OUTPUT
    uDays      : UDINT;                    (* 天分量，[d]，上界 24（TIME 容器毫秒上限 ÷ 86400）/ the days component, capped at 24 by the container *)
    uHours     : UDINT;                    (* 时分量，[h]，域 [0, 23] / the hours component, 0..23 *)
    uMins      : UDINT;                    (* 分分量，[min]，域 [0, 59] / the minutes component, 0..59 *)
    uSecs      : UDINT;                    (* 秒分量，[s]，域 [0, 59] / the seconds component, 0..59 *)
    bTruncated : BOOL;                     (* 毫秒余量非零被舍弃（显示口径向下取整到秒），[标志] / TRUE when a nonzero millisecond remainder was discarded *)
END_VAR
VAR CONSTANT
    DL_DUF_MS_DAY  : UDINT := 86400000;    (* 一天的毫秒数（常量除子，无变量除零面）/ the milliseconds per day, a constant divisor *)
    DL_DUF_MS_HOUR : UDINT := 3600000;     (* 一小时的毫秒数（常量除子）/ the milliseconds per hour, a constant divisor *)
    DL_DUF_MS_MIN  : UDINT := 60000;       (* 一分钟的毫秒数（常量除子）/ the milliseconds per minute, a constant divisor *)
    DL_DUF_MS_SEC  : UDINT := 1000;        (* 一秒的毫秒数（常量除子）/ the milliseconds per second, a constant divisor *)
END_VAR
VAR
    dMs   : DINT;                          (* 毫秒整数中间量（容器原值），[ms] / the millisecond integer temporary *)
    uMs   : UDINT;                         (* 毫秒无符号中间量，[ms] / the unsigned millisecond temporary *)
    uRem1 : UDINT;                         (* 天分解余数，[ms] / the remainder after the days split *)
    uRem2 : UDINT;                         (* 时分解余数，[ms] / the remainder after the hours split *)
    uRem3 : UDINT;                         (* 分分解余数，[ms] / the remainder after the minutes split *)
END_VAR

// 段 1｜返回值与分量预置（统一出口预置，R256）/ segment 1, preset the return and the components
FC_DL_DurationFormat := FALSE;             // 故障缺省返回不可信 / the fault default is not trustworthy
uDays      := 0;                           // 天分量预置零 / preset the days component to zero
uHours     := 0;                           // 时分量预置零 / preset the hours component to zero
uMins      := 0;                           // 分分量预置零 / preset the minutes component to zero
uSecs      := 0;                           // 秒分量预置零 / preset the seconds component to zero
bTruncated := FALSE;                       // 舍弃标志预清零 / preset the truncation flag false

// 段 2｜容器换算与负值防御闸（TIME 无符号语义，负值不可表示，防御性复检）/ segment 2, the container conversion and the negative guard
dMs := TIME_TO_DINT(tDur);                 // 容器毫秒原值（标准类型转换）/ the container value in ms, a standard conversion
IF dMs < 0 THEN                            // 负值不可表示（非法入参，防御兜底）/ a negative value is not representable
    RETURN;                                // 结构早退（分量保持清零预置，返回 FALSE）/ structural exit, the components stay zeroed
END_IF

// 段 3｜整除分解（常量除子级联，无变量除零面）/ segment 3, the integer division cascade
uMs   := DINT_TO_UDINT(dMs);               // 毫秒无符号化（已过负值闸，无负数面）/ the unsigned milliseconds, guarded
uDays := uMs / DL_DUF_MS_DAY;              // 天分量（整除向下取整）/ the days component
uRem1 := uMs MOD DL_DUF_MS_DAY;            // 天分解余数 / the remainder after days
uHours := uRem1 / DL_DUF_MS_HOUR;          // 时分量 / the hours component
uRem2 := uRem1 MOD DL_DUF_MS_HOUR;         // 时分解余数 / the remainder after hours
uMins := uRem2 / DL_DUF_MS_MIN;            // 分分量 / the minutes component
uRem3 := uRem2 MOD DL_DUF_MS_MIN;          // 分分解余数 / the remainder after minutes
uSecs := uRem3 / DL_DUF_MS_SEC;            // 秒分量 / the seconds component

// 段 4｜毫秒余量舍弃声明（bTruncated 名实对齐，边界四）/ segment 4, the millisecond remainder disclosure
bTruncated := (uRem3 MOD DL_DUF_MS_SEC) <> 0; // 余量非零即已舍弃 / a nonzero remainder was discarded

// 段 5｜正常出口 / segment 5, the normal outlet
FC_DL_DurationFormat := TRUE;              // 入参合法且已完整分解 / a valid input fully decomposed
END_FUNCTION

(* ---- FC_DL_DwordsToLword.st ---- *)
(*==============================================================================
 * 名称 : FC_DL_DwordsToLword —— 两个 DWORD 合成 LWORD（显式高低序参数）
 * 分类 / 前缀 / 版本 : DL_Base / FC_DL_ / 1.0.0
 * 溯源 : 开源语义参考（OSCAT/AixOCAT 族，MIT）或 clean-room IEC 实现，未复制源码
 * 平台 : 纯 IEC 61131-3
 * 功能说明 : 将两个 32 位 DWORD 合成为 64 位 LWORD：bFirstIsHigh=TRUE 时 dwFirst
 *            为高 32 位、dwSecond 为低 32 位；FALSE 时角色对调。
 *            合成全程数值语义（DWORD_TO_LWORD + SHL/OR），不触碰内存序。
 *            边界处理：两双字覆盖完整 64 位，无溢出；与 FC_DL_LwordToDwords
 *            互为逆运算（同参数口径下往返一致）。
 * 错误码 : 无故障路径（全值域合法的纯合成），eErr 恒 0，bValid 恒 TRUE；
 *          16#0001_1A0E 为本件预留码位，当前实现不发出
 * 状态机 : R6 标注 N/A（纯函数无顺序状态，以本节替代 ELSE 兜底）
 * 红线 : R1/R2/R3 ✓ 零全局/零IO/纯IEC ｜ R4 ✓ 移位量=32<64 ｜ R10 ✓ 标准转换 ｜ R11 ✓ 分号收尾 ｜ R15 ✓ 无保留字撞名
 * 修订记录 : 2026-11-23 v1.0.0 首次入库（R76）
 *============================================================================*)
FUNCTION FC_DL_DwordsToLword : LWORD
VAR_INPUT
    dwFirst     : DWORD;   // 首个输入双字 [位域] / first input dword
    dwSecond    : DWORD;   // 第二个输入双字 [位域] / second input dword
    bFirstIsHigh: BOOL;    // TRUE=dwFirst 为高 32 位 / TRUE when dwFirst is the high half
END_VAR
VAR_OUTPUT
    eErr   : UDINT;    // 故障码，0=正常（本件无故障路径）/ error code, 0=ok (no fault path)
    bError : BOOL;     // 故障标志，恒 FALSE / error flag, always FALSE
    bValid : BOOL;     // TRUE=返回值可用，恒 TRUE / TRUE when return value is usable
END_VAR
VAR
    _dwHi : DWORD;     // 判定后的高 32 位 / resolved high dword
    _dwLo : DWORD;     // 判定后的低 32 位 / resolved low dword
END_VAR

eErr   := 16#0000_0000;                      // 故障码清零 / clear error code
bError := FALSE;                             // 故障标志清零 / clear error flag
bValid := TRUE;                              // 本件全值域合法，恒可用 / always valid

IF bFirstIsHigh THEN                         // dwFirst 为高 32 位 / dwFirst is high
    _dwHi := dwFirst;                        // 取 dwFirst 为高 / take dwFirst as high
    _dwLo := dwSecond;                       // 取 dwSecond 为低 / take dwSecond as low
ELSE                                         // dwSecond 为高 32 位 / dwSecond is high
    _dwHi := dwSecond;                       // 取 dwSecond 为高 / take dwSecond as high
    _dwLo := dwFirst;                        // 取 dwFirst 为低 / take dwFirst as low
END_IF

FC_DL_DwordsToLword := SHL(DWORD_TO_LWORD(_dwHi), 32) OR DWORD_TO_LWORD(_dwLo);    // 高 32 位左移后并入低 32 位（移位量 32<64 安全）/ compose

END_FUNCTION

(* ---- FC_DL_DwordToWords.st ---- *)
(*==============================================================================
 * 名称 : FC_DL_DwordToWords —— DWORD 拆解为两个 WORD（本件返回首字，wOther 为次字）
 * 分类 / 前缀 / 版本 : DL_Base / FC_DL_ / 1.0.0
 * 溯源 : 开源语义参考（OSCAT/AixOCAT 族，MIT）或 clean-room IEC 实现，未复制源码
 * 平台 : 纯 IEC 61131-3
 * 功能说明 : 将 32 位输入拆为高/低两个 16 位 WORD。bHiFirst=TRUE 时首字（返回值）
 *            为高字、次字（wOther）为低字；FALSE 时角色对调（首字=低字）。
 *            「首/次」仅表拆解顺序，与内存字节序无关（数值语义拆解）。
 *            边界处理：dwIn 全值域合法，高低字覆盖完整 32 位，无信息丢失。
 * 错误码 : 无故障路径（全值域合法的纯拆解），eErr 恒 0，bValid 恒 TRUE；
 *          16#0001_1A0A 为本件预留码位，当前实现不发出
 * 状态机 : R6 标注 N/A（纯函数无顺序状态，以本节替代 ELSE 兜底）
 * 红线 : R1/R2/R3 ✓ 零全局/零IO/纯IEC ｜ R4 ✓ 移位量=16 ｜ R10 ✓ 标准转换 ｜ R11 ✓ 分号收尾 ｜ R15 ✓ 无保留字撞名
 * 修订记录 : 2026-11-23 v1.0.0 首次入库（R76）
 *============================================================================*)
FUNCTION FC_DL_DwordToWords : WORD
VAR_INPUT
    dwIn     : DWORD;    // 待拆解的 32 位输入 [位域] / input dword to be split
    bHiFirst : BOOL;     // TRUE=首字取高字 / TRUE when first word is the high word
END_VAR
VAR_OUTPUT
    wOther : WORD;     // 次字（另一半）/ the other (second) word
    eErr   : UDINT;    // 故障码，0=正常（本件无故障路径）/ error code, 0=ok (no fault path)
    bError : BOOL;     // 故障标志，恒 FALSE / error flag, always FALSE
    bValid : BOOL;     // TRUE=首/次两字均可用，恒 TRUE / TRUE when both words are usable
END_VAR
VAR
    _wHi : WORD;       // 高 16 位字 [位域] / high word
    _wLo : WORD;       // 低 16 位字 [位域] / low word
END_VAR

eErr   := 16#0000_0000;                      // 故障码清零 / clear error code
bError := FALSE;                             // 故障标志清零 / clear error flag
bValid := TRUE;                              // 本件全值域合法，恒可用 / always valid

_wHi := DWORD_TO_WORD(SHR(dwIn, 16));        // 右移 16 位取高字（截断安全）/ high word via shift
_wLo := DWORD_TO_WORD(dwIn AND 16#0000_FFFF);// 低 16 位掩码后截取 / low word via mask

IF bHiFirst THEN                             // 首字 = 高字 / first word is high word
    FC_DL_DwordToWords := _wHi;              // 返回首字为高字 / return high as first
    wOther := _wLo;                          // 次字为低字 / low as other
ELSE                                         // 首字 = 低字 / first word is low word
    FC_DL_DwordToWords := _wLo;              // 返回首字为低字 / return low as first
    wOther := _wHi;                          // 次字为高字 / high as other
END_IF

END_FUNCTION

(* ---- FC_DL_EndianProbe.st ---- *)
(*==============================================================================
 * 名称 : FC_DL_EndianProbe —— 运行期字节序探针（纯 IEC 语义层判定）
 * 分类 / 前缀 / 版本 : DL_Base / FC_DL_ / 1.0.0
 * 溯源 : 开源语义参考（OSCAT/AixOCAT 族，MIT）或 clean-room IEC 实现，未复制源码
 * 平台 : 纯 IEC 61131-3
 * 功能说明 : 返回 FALSE（判定为小端约定）且 bValid=TRUE。判定依据（非含糊占位）：
 *            (1) IEC 61131-3 第 3 版对 SHL/SHR/AND/OR 及 WORD_TO_BYTE 等转换的
 *                定义均在「数值语义」层，与目标机内存字节排布完全无关——把
 *                WORD 16#0102 经 SHR(...,8) 取出的是数值高字节 16#01，任何
 *                平台上该结论一致，故移位序列无法探测内存序；
 *            (2) R3 红线禁用 POINTER/REFERENCE/UNION，纯 IEC 层不存在合法的
 *                内存字节重解释手段，因此运行期探针在本库约束下不可实现；
 *            (3) 本库所有字节序件一律显式携带 bBigEndian/bHiFirst 参数、按
 *                数值语义装配/拆解，不依赖内存序，故探针恒判 FALSE（库级
 *                约定：小端数值语义），bValid 恒 TRUE 表示该约定全平台成立。
 * 错误码 : 无故障路径（常量语义判定），eErr 恒 0，bValid 恒 TRUE；
 *          16#0001_1A0C 为本件预留码位，当前实现不发出
 * 状态机 : R6 标注 N/A（纯函数无顺序状态，以本节替代 ELSE 兜底）
 * 红线 : R1/R2/R3 ✓ 零全局/零IO/纯IEC（禁指针/联合体）｜ R4 ✓ N/A 无浮点 ｜ R10 ✓ 标准转换 ｜ R11 ✓ 分号收尾 ｜ R15 ✓ 无保留字撞名
 * 修订记录 : 2026-11-23 v1.0.0 首次入库（R76）
 *============================================================================*)
FUNCTION FC_DL_EndianProbe : BOOL
VAR_OUTPUT
    eErr   : UDINT;    // 故障码，0=正常（本件无故障路径）/ error code, 0=ok (no fault path)
    bError : BOOL;     // 故障标志，恒 FALSE / error flag, always FALSE
    bValid : BOOL;     // TRUE=判定结论可用，恒 TRUE / TRUE when verdict is usable
END_VAR

eErr   := 16#0000_0000;                      // 故障码清零 / clear error code
bError := FALSE;                             // 故障标志清零 / clear error flag
bValid := TRUE;                              // 数值语义约定全平台成立 / verdict usable on all platforms

FC_DL_EndianProbe := FALSE;                  // 恒判 FALSE：库级小端数值语义约定 / always FALSE by library convention

END_FUNCTION
